// TIA Portal project "PalletWarehouse" (V20)

(* hardware
DEVICE "S7-1500/ET200MP-Station_1"  S7-1500 station
   slot 0: "Profilschiene_0"  Rack  6ES7 590-1***0-0AA0
   slot 1: "PLC_1"  CPU 1513-1 PN  6ES7 513-1AM03-0AB0  V4.0
      slot 3: "CPU-Display_1"  6ES7591-1AA00-0AA0
      slot 32768: "PROFINET-Schnittstelle_1"  X1
         slot 32769: "Port_1"  X1 P1
         slot 32770: "Port_2"  X1 P2
      slot 34817: "Virtual CP interface port_1"  Virtual CP interface port  Virtual CP interface port FW V4.0
   slot 2: "DI 16x24VDC BA_1"  DI 16x24VDC BA  6ES7 521-1BH10-0AA0  V1.1
   slot 3: "DQ 16x24VDC/0.5A ST_1"  DQ 16x24VDC/0.5A ST  6ES7 522-1BH00-0AB0  V2.0
   slot 4: "AI 8xU/I/R/RTD BA_1"  AI 8xU/I/R/RTD BA  6ES7 531-7QF00-0AB0  V1.0
   slot 5: "AQ 8xU/I HS_1"  AQ 8xU/I HS  6ES7 532-5HF00-0AB0  V2.2
   slot 6: "DQ 16x24VDC/0.5A ST_2"  DQ 16x24VDC/0.5A ST  6ES7 522-1BH00-0AB0  V2.0
   slot 7: "DI 16x24VDC BA_2"  DI 16x24VDC BA  6ES7 521-1BH10-0AA0  V1.1
   slot 8: "AQ 2xU/I ST_1"  AQ 2xU/I ST  6ES7 532-5NB00-0AB0  V1.0
   slot 9: "DI 16x24VDC BA_3"  DI 16x24VDC BA  6ES7 521-1BH10-0AA0  V1.1
DEVICE "PC-System_1"  SIMATIC PC station
   slot 0: "SIMATIC PC station"  Rail  SIMATIC PC-Station  V1.0
      slot 125: "Stationmanager"  Station_Manager  V6.0.4
   slot 1: "HMI_RT_1"  WinCC RT Advanced  6AV2 104-0xxxx-xxxx  17.0.0.0
      slot 33792: "Computer interface"  Host interface
   slot 2: "IE general_1"  IE General  IE_CP  V8.2.0
      slot 1: "PROFINET interface"  IEGeneral.Interface.8.2.0
*)

// ===== PLC "PLC_1"  CPU 1513-1 PN =====

VAR_GLOBAL   // PLC tag table "Standard-Variablentabelle"
   "PlcLabConnectIn01" AT %ID32760 : DWord;
   "PlcLabConnectIn02" AT %ID32764 : DWord;
   "PlcLabConnectOut01" AT %QD32760 : DWord;
   "PlcLabConnectOut02" AT %QD32764 : DWord;
END_VAR

VAR_GLOBAL   // PLC tag table "IO"
   "PalletizerEntrySensor" AT %I0.1 : Bool;
   "PusherLimitSensor" AT %I0.3 : Bool;
   "PalletizerBelt" AT %Q0.4 : Bool;
   "PalletizerTurn" AT %Q0.5 : Bool;
   "PusherMotor" AT %Q0.6 : Bool;
   "PalletizerClampedSensor" AT %I0.5 : Bool;
   "PalletizerPlateLimit" AT %I0.4 : Bool;
   "PalletizerElevatorMovingSensor" AT %I0.6 : Bool;
   "PalletizerClamp" AT %Q0.7 : Bool;
   "PalletizerPlate" AT %Q1.0 : Bool;
   "PalletizerElevatorUp" AT %Q1.1 : Bool;
   "PalletizerElevatorDown" AT %Q1.2 : Bool;
   "PalletizerElevatorMoveToLimit" AT %Q1.3 : Bool;
   "BoxEmitter" AT %Q0.1 : Bool;
   "PalletChainFrontLimit" AT %I0.7 : Bool;
   "BoxFeedConveyor" AT %Q0.0 : Bool;
   "PalletChain" AT %Q0.2 : Bool;
   "PalletFeedSensor" AT %I0.2 : Bool;
   "PalletFeedConveyor" AT %Q1.4 : Bool;
   "PalletEmitter" AT %Q0.3 : Bool;
   "ConveyorSensor1" AT %I1.1 : Bool;
   "ConveyorSensor2" AT %I1.2 : Bool;
   "TransferConveyor1" AT %Q1.5 : Bool;
   "TransferConveyor2" AT %Q1.6 : Bool;
   "TurntableEntrySensor" AT %I1.3 : Bool;
   "PalletChainBackLimit" AT %I1.0 : Bool;
   "TurntableTurn" AT %Q1.7 : Bool;
   "TurntableRollForward" AT %Q2.0 : Bool;
   "TurntableRollBackward" AT %Q2.1 : Bool;
   "TurntableLimit0" AT %I1.4 : Bool;
   "TurntableLimit90" AT %I1.5 : Bool;
   "TurntableBackLimit" AT %I1.6 : Bool;
   "TurntableFrontLimit" AT %I1.7 : Bool;
   "TurntableLeftExitSensor" AT %I2.0 : Bool;
   "TurntableRightExitSensor" AT %I2.1 : Bool;
   "Crane1MovingX" AT %I2.2 : Bool;
   "Crane1MovingZ" AT %I2.3 : Bool;
   "Crane1LeftLimit" AT %I2.4 : Bool;
   "Crane1RightLimit" AT %I2.5 : Bool;
   "Crane1Lift" AT %Q2.2 : Bool;
   "Crane1Right" AT %Q2.4 : Bool;
   "Crane1Left" AT %Q2.3 : Bool;
   "Crane1Position" AT %QW30 : Int;
   "StartButtonTemp" AT %I2.7 : Bool;
   "Crane1MidLimit" AT %I2.6 : Bool;
   "Crane2MovingX" AT %I3.0 : Bool;
   "Crane2MovingZ" AT %I3.1 : Bool;
   "Crane2LeftLimit" AT %I3.2 : Bool;
   "Crane2RightLimit" AT %I3.3 : Bool;
   "Crane2MidLimit" AT %I3.4 : Bool;
   "Crane2Lift" AT %Q2.5 : Bool;
   "Crane2Right" AT %Q2.7 : Bool;
   "Crane2Left" AT %Q2.6 : Bool;
   "Crane2Position" AT %QW32 : Int;
   "LoadSensor1" AT %I3.5 : Bool;
   "LoadSensor2" AT %I3.6 : Bool;
   "LoadConveyor1" AT %Q3.0 : Bool;
   "LoadConveyor2" AT %Q3.1 : Bool;
   "BoxEmitterSensor" AT %I0.0 : Bool;
   "UnloadSensor1" AT %I3.7 : Bool;
   "UnloadSensor2" AT %I4.0 : Bool;
   "RemoverSensor1" AT %I4.1 : Bool;
   "RemoverSensor2" AT %I4.2 : Bool;
   "UnloadConveyor1" AT %Q3.2 : Bool;
   "UnloadConveyor2" AT %Q3.3 : Bool;
   "RemoverConveyor1" AT %Q3.4 : Bool;
   "RemoverConveyor2" AT %Q3.5 : Bool;
   "Remover1" AT %Q3.6 : Bool;
   "Remover2" AT %Q3.7 : Bool;
END_VAR

TYPE "StorageCraneUDT"
   STRUCT
      CraneSides : Struct
         LoadRight : Bool;
         UnloadRight : Bool;
         PickupRight : Bool;
      END_STRUCT;
      In : Struct
         MovingX : Bool;
         MovingZ : Bool;
         LeftLimit : Bool;
         RightLimit : Bool;
         MidLimit : Bool;
      END_STRUCT;
      Out : Struct
         Lift : Bool;
         Left : Bool;
         Right : Bool;
         Position : Int;
      END_STRUCT;
   END_STRUCT;
END_TYPE

TYPE "WarehouseSlotUDT"
   STRUCT
      Id : Int;
      Status : Int;
      "Time" : DTL;
   END_STRUCT;
END_TYPE

TYPE "PalletizerUDT"
   STRUCT
      In : Struct
         BoxEntrySensor : Bool;
         PusherLimit : Bool;
         Clamped : Bool;
         PlateLimit : Bool;
         ElevatorMoving : Bool;
         ElevatorFrontLimit : Bool;
         ElevatorBackLimit : Bool;
         PalletFeedSensor : Bool;
         EmitSensor : Bool;
      END_STRUCT;
      Out : Struct
         PalletFeedConv : Bool;
         BoxFeedConv : Bool;
         Turn : Bool;
         Clamp : Bool;
         Pusher : Bool;
         Plate : Bool;
         ElevatorUp : Bool;
         ElevatorDown : Bool;
         ElevatorMoveToLimit : Bool;
         PalletConv : Bool;
         PalletEmitter : Bool;
         EmitConv : Bool;
         BoxEmitter : Bool;
      END_STRUCT;
   END_STRUCT;
END_TYPE

TYPE "ConveyorUDT"
   STRUCT
      In : Struct
         StartSensor : Bool;
         EndSensor : Bool;
         Stop : Bool;
      END_STRUCT;
      Out : Struct
         Conveyor : Bool;
      END_STRUCT;
   END_STRUCT;
END_TYPE

TYPE "TurntableUDT"
   STRUCT
      In : Struct
         FrontLimit : Bool;
         BackLimit : Bool;
         Limit90 : Bool;
         Limit0 : Bool;
      END_STRUCT;
      Out : Struct
         RollForward : Bool;
         RollBackward : Bool;
         Turn : Bool;
      END_STRUCT;
   END_STRUCT;
END_TYPE

DATA_BLOCK "Warehouse_DB"   // DB9
{ S7_Optimized_Access := 'TRUE' }
VERSION : 0.1
// stored: InstanceOfName Warehouse
"Warehouse"
BEGIN
END_DATA_BLOCK

// folder: HMI

DATA_BLOCK "HMI_Data"   // DB11
{ S7_Optimized_Access := 'TRUE' }
VERSION : 0.1
   VAR
      SelectedRack : Int;
      SelectedSlot : Int;
      TargetSlot : "WarehouseSlotUDT";
      RetrievePallet : Bool;
      StopCmd : Bool;
      StartCmd : Bool;
      RacksFull : Bool;
      CraneStatus : Array[1..2] of Int;
      OccupiedSlots : Array[1..2] of Int;
   END_VAR
BEGIN
END_DATA_BLOCK

// folder: IO Mapping

DATA_BLOCK "IO"   // DB2
{ S7_Optimized_Access := 'TRUE' }
VERSION : 0.1
   VAR
      Palletizer : "PalletizerUDT";
      StorageCrane1 : "StorageCraneUDT";
      StorageCrane2 : "StorageCraneUDT";
      LineIO : Struct
         TransferConveyor1IO : "ConveyorUDT";
         TransferConveyor2IO : "ConveyorUDT";
         LoadConveyor1IO : "ConveyorUDT";
         LoadConveyor2IO : "ConveyorUDT";
         UnloadConveyor1IO : "ConveyorUDT";
         UnloadConveyor2IO : "ConveyorUDT";
         TurntableIO : "TurntableUDT";
         Remover1 : Bool;
         Remover2 : Bool;
      END_STRUCT;
   END_VAR
BEGIN
   StorageCrane1.CraneSides.LoadRight := TRUE;
   StorageCrane1.CraneSides.PickupRight := TRUE;
   StorageCrane1.CraneSides.UnloadRight := FALSE;
   StorageCrane2.CraneSides.PickupRight := FALSE;
   StorageCrane2.CraneSides.UnloadRight := TRUE;
   StorageCrane2.CraneSides.LoadRight := TRUE;
END_DATA_BLOCK

// folder: WarehouseManager

DATA_BLOCK "WarehouseData"   // DB10
{ S7_Optimized_Access := 'TRUE' }
VERSION : 0.1
   VAR
      Rack1 : Array[1..54] of "WarehouseSlotUDT";
      Rack2 : Array[1..54] of "WarehouseSlotUDT";
   END_VAR
BEGIN
END_DATA_BLOCK

// folder: (top level)

FUNCTION_BLOCK "Warehouse"   // FB15, SCL
{ S7_Optimized_Access := 'TRUE' }
VERSION : 0.1
   VAR_IN_OUT
      PalletizerIO : "PalletizerUDT";
      StorageCrane1IO : "StorageCraneUDT";
      StorageCrane2IO : "StorageCraneUDT";
      LineIO : Struct
         TransferConveyor1IO : "ConveyorUDT";
         TransferConveyor2IO : "ConveyorUDT";
         LoadConveyor1IO : "ConveyorUDT";
         LoadConveyor2IO : "ConveyorUDT";
         UnloadConveyor1IO : "ConveyorUDT";
         UnloadConveyor2IO : "ConveyorUDT";
         TurntableIO : "TurntableUDT";
         Remover1 : Bool;
         Remover2 : Bool;
      END_STRUCT;
   END_VAR
   VAR
      Line : "Line";
      WarehouseManager : "WarehouseManager";
      CraneLoadDone : Array[1..2] of Bool;
      CraneUnloadDone : Array[1..2] of Bool;
      CraneBusy : Array[1..2] of Bool;
      Palletizer : "Palletizer";
      StorageCrane1 : "StorageCrane";
      StorageCrane2 : "StorageCrane";
      WarehouseControl : "WarehouseControl";
   END_VAR
BEGIN
   #WarehouseControl(StartCmd := "HMI_Data".StartCmd,
                     StopCmd := "HMI_Data".StopCmd,
                     Active := false);

   #Palletizer(PalletizerIO:=#PalletizerIO,
               Run:=#WarehouseControl.Run AND NOT #WarehouseManager.Full);

   #WarehouseManager(UnloadDone:=#CraneUnloadDone,
                     CraneBusy:=#CraneBusy,
                     PalletReady := #LineIO.TransferConveyor2IO.In.EndSensor,
                     UnloadRequest:="HMI_Data".RetrievePallet,
                     UnloadRack:="HMI_Data".SelectedRack,
                     UnloadSlot:="HMI_Data".SelectedSlot,
                     Run:=#WarehouseControl.Run,
                     Rack1Slots := "WarehouseData".Rack1,
                     Rack2Slots := "WarehouseData".Rack2,
                     LoadDone:=#CraneLoadDone,
                     Full=>"HMI_Data".RacksFull,
                     CraneStatus=>"HMI_Data".CraneStatus); 

   #Line(TurntableRollDirection:=#WarehouseManager.Rack,
         Run:=#WarehouseControl.Run,
         Remover1=>#LineIO.Remover1,
         Remover2=>#LineIO.Remover2,
         TransferConveyor1IO:=#LineIO.TransferConveyor1IO,
         TransferConveyor2IO:=#LineIO.TransferConveyor2IO,
         LoadConveyor1IO:=#LineIO.LoadConveyor1IO,
         LoadConveyor2IO:=#LineIO.LoadConveyor2IO,
         UnloadConveyor1IO:=#LineIO.UnloadConveyor1IO,
         UnloadConveyor2IO:=#LineIO.UnloadConveyor2IO,
         TurntableIO:=#LineIO.TurntableIO);

   #StorageCrane1(TargetPosition:=#WarehouseManager.TargetSlot[1],
                  RequestLoad:=#WarehouseManager.LoadStart[1] AND #LineIO.LoadConveyor1IO.In.Stop,
                  RequestUnload:=#WarehouseManager.UnloadStart[1],
                  Run:=#WarehouseControl.Run,
                  LoadDone=>#CraneLoadDone[1],
                  UnloadDone=>#CraneUnloadDone[1],
                  StorageCraneUDT:=#StorageCrane1IO,
                  Busy=>#CraneBusy[1]); 

   #StorageCrane2(TargetPosition := #WarehouseManager.TargetSlot[2],
                  RequestLoad := #WarehouseManager.LoadStart[2] AND #LineIO.LoadConveyor2IO.In.Stop,
                  RequestUnload := #WarehouseManager.UnloadStart[2],
                  Run:=#WarehouseControl.Run,
                  LoadDone => #CraneLoadDone[2],
                  UnloadDone=>#CraneUnloadDone[2],
                  StorageCraneUDT := #StorageCrane2IO,
                  Busy=>#CraneBusy[2]);
END_FUNCTION_BLOCK

FUNCTION_BLOCK "WarehouseControl"   // FB19, SCL
{ S7_Optimized_Access := 'TRUE' }
VERSION : 0.1
   VAR_INPUT
      StartCmd : Bool;
      StopCmd : Bool;
      Active : Bool;
   END_VAR
   VAR_OUTPUT
      Run : Bool;
      Status : Int;
   END_VAR
   VAR
      StopPEdge : R_TRIG;
      StartPEdge : R_TRIG;
   END_VAR
BEGIN
   #StartPEdge(CLK:=#StartCmd);
   #StopPEdge(CLK := #StopCmd);

   IF #StopPEdge.Q THEN
       #Run := FALSE;
   ELSIF #StartPEdge.Q THEN
       #Run := TRUE;
   END_IF;

   IF #Run THEN
       #Status := 1;
   ELSIF #Active THEN
       #Status := 2;
   ELSE
       #Status := 0;
   END_IF;
END_FUNCTION_BLOCK

ORGANIZATION_BLOCK "Main"   // OB1, LAD, ProgramCycle
TITLE = "Main Program Sweep (Cycle)"
{ S7_Optimized_Access := 'TRUE' }
VERSION : 0.1
   VAR_INPUT
      Initial_Call : Bool;   // Initial call of this OB
      Remanence : Bool;   // =True, if remanent data are available
   END_VAR
BEGIN

REGION Network 1
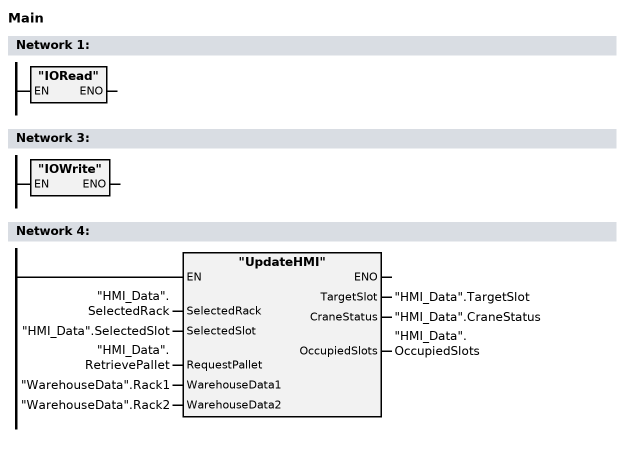
   RUNG wire#powerrail
      "IORead"()
   END_RUNG
   // the same network as SCL:
   "IORead"();
END_REGION

REGION Network 2 (SCL)
   "Warehouse_DB"(PalletizerIO:="IO".Palletizer,
                  StorageCrane1IO:="IO".StorageCrane1,
                  StorageCrane2IO:="IO".StorageCrane2,
                  LineIO:="IO".LineIO);
END_REGION

REGION Network 3
   RUNG wire#powerrail
      "IOWrite"()
   END_RUNG
   // the same network as SCL:
   "IOWrite"();
END_REGION

REGION Network 4
   RUNG wire#powerrail
      "UpdateHMI"(SelectedRack := "HMI_Data".SelectedRack, SelectedSlot := "HMI_Data".SelectedSlot, RequestPallet := "HMI_Data".RetrievePallet, WarehouseData1 := "WarehouseData".Rack1, WarehouseData2 := "WarehouseData".Rack2, TargetSlot => "HMI_Data".TargetSlot, CraneStatus => "HMI_Data".CraneStatus, OccupiedSlots => "HMI_Data".OccupiedSlots)
   END_RUNG
   // the same network as SCL:
   "UpdateHMI"(SelectedRack := "HMI_Data".SelectedRack,
               SelectedSlot := "HMI_Data".SelectedSlot,
               RequestPallet := "HMI_Data".RetrievePallet,
               WarehouseData1 := "WarehouseData".Rack1,
               WarehouseData2 := "WarehouseData".Rack2,
               TargetSlot => "HMI_Data".TargetSlot,
               CraneStatus => "HMI_Data".CraneStatus,
               OccupiedSlots => "HMI_Data".OccupiedSlots);
END_REGION
END_ORGANIZATION_BLOCK

// folder: HMI

FUNCTION "UpdateHMI" : Void   // FC6, SCL
{ S7_Optimized_Access := 'TRUE' }
VERSION : 0.1
   VAR_INPUT
      SelectedRack : Int;
      SelectedSlot : Int;
      RequestPallet : Bool;
      WarehouseData1 : Array[1..54] of "WarehouseSlotUDT";
      WarehouseData2 : Array[1..54] of "WarehouseSlotUDT";
   END_VAR
   VAR_OUTPUT
      TargetSlot : "WarehouseSlotUDT";
      CraneStatus : Array[1..2] of Int;
      OccupiedSlots : Array[1..2] of Int;
   END_VAR
   VAR_TEMP
      i : Int;
      freeslots : Array[1..2] of Int;
   END_VAR
BEGIN
   IF #SelectedRack = 1 THEN
       #TargetSlot := #WarehouseData1[#SelectedSlot];
   ELSIF #SelectedRack = 2 THEN
       #TargetSlot := #WarehouseData2[#SelectedSlot];
   END_IF;

   #freeslots[1]:="CountFreeSlots"(#WarehouseData1);
   #freeslots[2] := "CountFreeSlots"(#WarehouseData2);

   FOR #i := 1 TO 2 DO
       #OccupiedSlots[#i] := 54 - #freeslots[#i];
   END_FOR;
END_FUNCTION

// folder: IO Mapping

FUNCTION "IOWrite" : Void   // FC4, SCL
{ S7_Optimized_Access := 'TRUE' }
VERSION : 0.1
BEGIN
   // Mapping palletizer outputs
   "PalletFeedConveyor":="IO".Palletizer.Out.PalletFeedConv;
   "PalletizerBelt" :="IO".Palletizer.Out.BoxFeedConv;
   "PalletizerTurn" :="IO".Palletizer.Out.Turn;
   "PalletizerClamp":="IO".Palletizer.Out.Clamp;
   "PusherMotor" :="IO".Palletizer.Out.Pusher;
   "PalletizerPlate" := "IO".Palletizer.Out.Plate;
   "PalletizerElevatorUp" := "IO".Palletizer.Out.ElevatorUp;
   "PalletizerElevatorDown" :="IO".Palletizer.Out.ElevatorDown;
   "PalletizerElevatorMoveToLimit" :="IO".Palletizer.Out.ElevatorMoveToLimit;
   "PalletChain":="IO".Palletizer.Out.PalletConv;
   "PalletEmitter":="IO".Palletizer.Out.PalletEmitter;
   "BoxEmitter" := "IO".Palletizer.Out.BoxEmitter;
   "BoxFeedConveyor" := "IO".Palletizer.Out.EmitConv;

   // Mapping storage crane 1 outputs
   "Crane1Lift" := "IO".StorageCrane1.Out.Lift;
   "Crane1Left" :="IO".StorageCrane1.Out.Left;
   "Crane1Right" := "IO".StorageCrane1.Out.Right;
   "Crane1Position" := "IO".StorageCrane1.Out.Position;
   // Mapping storage crane 2 outputs
   "Crane2Lift":="IO".StorageCrane2.Out.Lift;
   "Crane2Left":="IO".StorageCrane2.Out.Left;
   "Crane2Right":="IO".StorageCrane2.Out.Right;
   "Crane2Position" := "IO".StorageCrane2.Out.Position;
   // Mapping line outputs
   "TransferConveyor1":="IO".LineIO.TransferConveyor1IO.Out.Conveyor;
   "TransferConveyor2":="IO".LineIO.TransferConveyor2IO.Out.Conveyor;
   "TurntableRollForward" := "IO".LineIO.TurntableIO.Out.RollForward;
   "TurntableRollBackward" := "IO".LineIO.TurntableIO.Out.RollBackward;
   "TurntableTurn" := "IO".LineIO.TurntableIO.Out.Turn;
   "LoadConveyor1":="IO".LineIO.LoadConveyor1IO.Out.Conveyor;
   "LoadConveyor2":="IO".LineIO.LoadConveyor2IO.Out.Conveyor;
   "UnloadConveyor1" := "IO".LineIO.UnloadConveyor1IO.Out.Conveyor;
   "UnloadConveyor2" := "IO".LineIO.UnloadConveyor2IO.Out.Conveyor;
   "RemoverConveyor1" := "IO".LineIO.UnloadConveyor1IO.Out.Conveyor;
   "RemoverConveyor2" := "IO".LineIO.UnloadConveyor2IO.Out.Conveyor;
   "Remover1" := "IO".LineIO.Remover1;
   "Remover2" := "IO".LineIO.Remover2;
END_FUNCTION

FUNCTION "IORead" : Void   // FC5, SCL
{ S7_Optimized_Access := 'TRUE' }
VERSION : 0.1
BEGIN
   // Mapping Palletizer Inputs
   "IO".Palletizer.In.BoxEntrySensor := "PalletizerEntrySensor";
   "IO".Palletizer.In.PusherLimit := "PusherLimitSensor";
   "IO".Palletizer.In.Clamped := "PalletizerClampedSensor";
   "IO".Palletizer.In.PlateLimit := "PalletizerPlateLimit";
   "IO".Palletizer.In.ElevatorMoving := "PalletizerElevatorMovingSensor";
   "IO".Palletizer.In.ElevatorFrontLimit := "PalletChainFrontLimit";
   "IO".Palletizer.In.ElevatorBackLimit := "PalletChainBackLimit";
   "IO".Palletizer.In.PalletFeedSensor := "PalletFeedSensor";
   "IO".Palletizer.In.EmitSensor := "BoxEmitterSensor";
   // Maping Storage Crane 1 Inputs
   "IO".StorageCrane1.In.MovingX := "Crane1MovingX";
   "IO".StorageCrane1.In.MovingZ := "Crane1MovingZ";
   "IO".StorageCrane1.In.LeftLimit := "Crane1LeftLimit";
   "IO".StorageCrane1.In.RightLimit := "Crane1RightLimit";
   "IO".StorageCrane1.In.MidLimit := "Crane1MidLimit";
   // Maping Storage Crane 2 Inputs
   "IO".StorageCrane2.In.MovingX := "Crane2MovingX";
   "IO".StorageCrane2.In.MovingZ := "Crane2MovingZ";
   "IO".StorageCrane2.In.LeftLimit := "Crane2LeftLimit";
   "IO".StorageCrane2.In.RightLimit := "Crane2RightLimit";
   "IO".StorageCrane2.In.MidLimit := "Crane2MidLimit";
   // Maping Line Inputs
   "IO".LineIO.TransferConveyor1IO.In.StartSensor := "ConveyorSensor1";
   "IO".LineIO.TransferConveyor1IO.In.EndSensor := "ConveyorSensor2";
   "IO".LineIO.TransferConveyor2IO.In.StartSensor := "ConveyorSensor2";
   "IO".LineIO.TransferConveyor2IO.In.EndSensor := "TurntableEntrySensor";
   "IO".LineIO.TurntableIO.In.FrontLimit := "TurntableFrontLimit";
   "IO".LineIO.TurntableIO.In.BackLimit := "TurntableBackLimit";
   "IO".LineIO.TurntableIO.In.Limit90 := "TurntableLimit90";
   "IO".LineIO.TurntableIO.In.Limit0 := "TurntableLimit0";
   "IO".LineIO.LoadConveyor1IO.In.StartSensor := "TurntableLeftExitSensor";
   "IO".LineIO.LoadConveyor1IO.In.Stop := "LoadSensor1";
   "IO".LineIO.LoadConveyor2IO.In.StartSensor := "TurntableRightExitSensor";
   "IO".LineIO.LoadConveyor2IO.In.Stop := "LoadSensor2";
   "IO".LineIO.UnloadConveyor1IO.In.StartSensor := "UnloadSensor1";
   "IO".LineIO.UnloadConveyor2IO.In.StartSensor := "UnloadSensor2";
   "IO".LineIO.UnloadConveyor1IO.In.Stop := "RemoverSensor1";
   "IO".LineIO.UnloadConveyor2IO.In.Stop := "RemoverSensor2";
END_FUNCTION

// folder: Line

FUNCTION_BLOCK "Line"   // FB1, LAD
{ S7_Optimized_Access := 'TRUE' }
VERSION : 0.1
   VAR_INPUT
      TurntableRollDirection : Int;
      Run : Bool;
   END_VAR
   VAR_OUTPUT
      Remover1 : Bool;
      Remover2 : Bool;
   END_VAR
   VAR_IN_OUT
      TransferConveyor1IO : "ConveyorUDT";
      TransferConveyor2IO : "ConveyorUDT";
      LoadConveyor1IO : "ConveyorUDT";
      LoadConveyor2IO : "ConveyorUDT";
      UnloadConveyor1IO : "ConveyorUDT";
      UnloadConveyor2IO : "ConveyorUDT";
      TurntableIO : "TurntableUDT";
   END_VAR
   VAR
      UnloadConveyor2 : "Conveyor";
      TransferConveyor1 : "Conveyor";
      TransferConveyor2 : "Conveyor";
      Turntable : "Turntable";
      LoadConveyor1 : "Conveyor";
      LoadConveyor2 : "Conveyor";
      UnloadConveyor1 : "Conveyor";
   END_VAR
BEGIN

REGION Network 1 (SCL)
   #TransferConveyor1(NextFree:=NOT #TransferConveyor2.Busy,
                      Run:=#Run,
                      ConveyorIO:=#TransferConveyor1IO);  

   #TransferConveyor2(NextFree:=TRUE,
                      Run:=#Run,
                      ConveyorIO:=#TransferConveyor2IO);

   #Turntable(Start:=#TransferConveyor2IO.In.EndSensor,
              Run:=#Run,
              RollDirection:=#TurntableRollDirection,
              RightSensor:=#LoadConveyor2IO.In.StartSensor,
              LeftSensor:=#LoadConveyor1IO.In.StartSensor,
              TurntableIO:=#TurntableIO); 

   #LoadConveyor1(NextFree:=TRUE,
                  Run:=#Run,
                  ConveyorIO:=#LoadConveyor1IO);

   #LoadConveyor2(NextFree:=TRUE,
                  Run:=#Run,
                  ConveyorIO:=#LoadConveyor2IO);

   #UnloadConveyor1(NextFree:=TRUE,
                    Run:=#Run,
                    ConveyorIO:=#UnloadConveyor1IO);

   #UnloadConveyor2(NextFree:=TRUE,
                    Run:=#Run,
                    ConveyorIO:=#UnloadConveyor2IO);

   #Remover1 := #UnloadConveyor1IO.In.Stop;
   #Remover2 := #UnloadConveyor2IO.In.Stop;
END_REGION
END_FUNCTION_BLOCK

FUNCTION_BLOCK "Conveyor"   // FB2, LAD
{ S7_Optimized_Access := 'TRUE' }
VERSION : 0.1
   VAR_INPUT
      NextFree : Bool;
      Run : Bool;
   END_VAR
   VAR_OUTPUT
      Busy : Bool;
   END_VAR
   VAR_IN_OUT
      ConveyorIO : "ConveyorUDT";
   END_VAR
   VAR
      Reset : Bool;
      Timeout_Instance : TON_TIME;
      Timeout : Bool;
      StartSensorEdge : Bool;
      EndSensorEdge : Bool;
      ConveyorStart : Bool;
   END_VAR
   VAR_TEMP   // added for the SCL form of the ladder/FBD networks
      _w1 : Bool;
   END_VAR
BEGIN

REGION Network 1
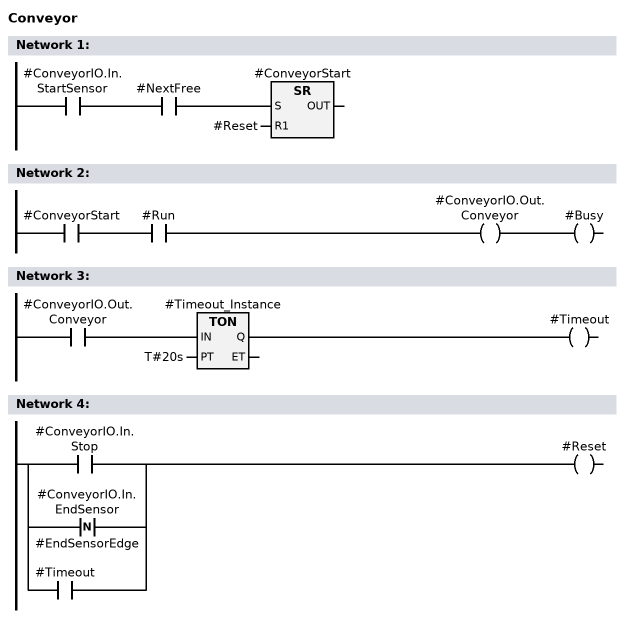
   RUNG wire#powerrail
      Contact( #ConveyorIO.In.StartSensor )
      Contact( #NextFree )
      S_SR(operand := #ConveyorStart, r1 := #Reset)
   END_RUNG
   // the same network as SCL:
   IF #ConveyorIO.In.StartSensor AND #NextFree THEN
       #ConveyorStart := TRUE;   // SR flip-flop
   END_IF;
   IF #Reset THEN #ConveyorStart := FALSE; END_IF;
END_REGION

REGION Network 2
   RUNG wire#powerrail
      Contact( #ConveyorStart )
      Contact( #Run )
      Coil( #ConveyorIO.Out.Conveyor )
      Coil( #Busy )
   END_RUNG
   // the same network as SCL:
   #ConveyorIO.Out.Conveyor := #ConveyorStart AND #Run;
   #Busy := #ConveyorIO.Out.Conveyor;
END_REGION

REGION Network 3
   #Timeout_Instance(IN := #ConveyorIO.Out.Conveyor, PT := T#20s);   // TON
   #Timeout := #Timeout_Instance.Q;
END_REGION

REGION Network 4
   RUNG wire#powerrail
      Contact( #ConveyorIO.In.Stop )
      wire#w1
      Coil( #Reset )
   END_RUNG
   RUNG wire#powerrail
      N_Contact(operand := #ConveyorIO.In.EndSensor, bit := #EndSensorEdge)
   END_RUNG wire#w1
   RUNG wire#powerrail
      Contact( #Timeout )
   END_RUNG wire#w1
   // the same network as SCL:
   #_w1 := NOT #ConveyorIO.In.EndSensor AND #EndSensorEdge;   // falling edge of #ConveyorIO.In.EndSensor
   #EndSensorEdge := #ConveyorIO.In.EndSensor;
   #Reset := #ConveyorIO.In.Stop OR #_w1 OR #Timeout;
END_REGION
END_FUNCTION_BLOCK

FUNCTION_BLOCK "Turntable"   // FB7, SCL
{ S7_Optimized_Access := 'TRUE' }
VERSION : 0.1
   VAR_INPUT
      Start : Bool;
      Run : Bool;
      RollDirection : Int;
      RightSensor : Bool;
      LeftSensor : Bool;
   END_VAR
   VAR_IN_OUT
      TurntableIO : "TurntableUDT";
   END_VAR
   VAR
      State : Int := 1;
      RightSensorNEdge : F_TRIG;
      LeftSensorNEdge : F_TRIG;
   END_VAR
BEGIN
   #RightSensorNEdge(CLK:=#RightSensor);
   #LeftSensorNEdge(CLK:=#LeftSensor);

   CASE #State OF
       1:  // Init
           IF #Start THEN
               #State := 2;
           END_IF;
           ;
       2:  // Load
           "IO".LineIO.TurntableIO.Out.RollForward := #Run;
           IF #TurntableIO.In.FrontLimit THEN
               #TurntableIO.Out.RollForward := FALSE;
               #State := 3;
           END_IF;
           ;
       3: // Turn
           #TurntableIO.Out.Turn := TRUE;
           IF #TurntableIO.In.Limit90 THEN
               #State := 4;
           END_IF;
       4: // Direction
           IF #RollDirection=1 THEN
               #State := 5;
           ELSIF #RollDirection=2 THEN
               #State := 6;
           END_IF;
       5: // Roll left
           #TurntableIO.Out.RollForward := #Run;
           IF #LeftSensorNEdge.Q THEN
               #TurntableIO.Out.RollForward := FALSE;
               #State := 7;
           END_IF;
       6: // Roll right
           #TurntableIO.Out.RollBackward := #Run;
           IF #RightSensorNEdge.Q THEN
               #TurntableIO.Out.RollBackward := FALSE;
               #State := 7;
           END_IF;
       7: // Return 
           #TurntableIO.Out.Turn := FALSE;
           IF #TurntableIO.In.Limit0 THEN
               #State := 1;
           END_IF;
   END_CASE;
END_FUNCTION_BLOCK

// folder: Palletizer

FUNCTION_BLOCK "Palletizer"   // FB3, SCL
{ S7_Optimized_Access := 'TRUE' }
VERSION : 0.1
   VAR_INPUT
      Run : Bool;
   END_VAR
   VAR_OUTPUT
      Busy : Bool;
   END_VAR
   VAR_IN_OUT
      PalletizerIO : "PalletizerUDT";
   END_VAR
   VAR
      State : Int := 1;
      BoxCount : Int := 0;
      BoxFeedTimer : TON_TIME;
      BoxFeedBusy : Bool;
      StackVertical : Bool := TRUE;
      PushCount : Int;
      BoxEntrySensorNEdge : F_TRIG;
      PusherFB : "Cylinder";
      BoxPerPush : Int;
      PushPerLayer : Int;
      PlateFB : "Cylinder";
      ElevatorFB : "Elevator";
      LayerCount : Int;
      PalletFeederFB : "PalletFeeder";
      BoxFeeder : "BoxFeedConv";
      UnloadConv : Bool;
   END_VAR
BEGIN
   #BoxEntrySensorNEdge(CLK := #PalletizerIO.In.BoxEntrySensor);
   #BoxFeedTimer(IN:=#PalletizerIO.Out.BoxFeedConv AND #BoxCount=#BoxPerPush,
                 PT:=T#2s);

   #PusherFB.Extend := FALSE;
   #PlateFB.Extend := FALSE;
   #PalletizerIO.Out.Clamp := FALSE;
   #PalletizerIO.Out.PalletConv := FALSE;
   #PalletFeederFB.Start := FALSE;
   #ElevatorFB.RequestUp := FALSE;
   #ElevatorFB.RequestDown := FALSE;
   #ElevatorFB.GoToLimit := FALSE;
   #UnloadConv := FALSE;

   IF #BoxEntrySensorNEdge.Q THEN
       #BoxCount := #BoxCount + 1;
   END_IF;

   IF #StackVertical THEN
       #PalletizerIO.Out.Turn := FALSE;
       #BoxPerPush := 2;
       #PushPerLayer := 3;
   ELSE
       #PalletizerIO.Out.Turn := TRUE;
       #BoxPerPush := 3;
       #PushPerLayer := 2;
   END_IF;

   CASE #State OF
       1:  // Init
           #StackVertical := True;
           #PushCount := 0;
           #BoxCount := 0;
           #LayerCount := 0;
           IF #Run THEN
               #State := 2;
           END_IF;
       2: // Pallet feed
           #PalletFeederFB.Start := #Run;
           IF #PalletFeederFB.Done THEN
               #State := 3;
           END_IF;

       3: // Elevator ready
           #ElevatorFB.GoToLimit := TRUE;
           #ElevatorFB.RequestUp := TRUE;
           IF #ElevatorFB.Done THEN
               #State := 4;
           END_IF;

       4:  // Box feed
           IF #PalletizerIO.In.BoxEntrySensor AND (#BoxCount < #BoxPerPush) AND #Run THEN
               #PalletizerIO.Out.BoxFeedConv := TRUE;
           ELSIF #BoxFeedTimer.Q THEN
               #PalletizerIO.Out.BoxFeedConv := FALSE;
           ELSIF (#BoxCount<#BoxPerPush) AND (NOT #Run) THEN
               #PalletizerIO.Out.BoxFeedConv := FALSE;
           END_IF;

           IF #BoxCount = #BoxPerPush AND NOT #PalletizerIO.Out.BoxFeedConv THEN
               #BoxCount := 0;
               #State := 5;
           END_IF;

       5:  // Extend pusher
           #PusherFB.Extend := TRUE;
           IF #PusherFB.Extended THEN
               #PushCount := #PushCount + 1;
               #State := 6;
           END_IF;

       6:  // Retract pusher
           IF #PusherFB.Retracted THEN
               IF #PushCount >= #PushPerLayer THEN
                   #PushCount := 0;
                   #StackVertical := NOT #StackVertical;
                   #State := 7;
               ELSE
                   #State := 4;
               END_IF;
           END_IF;

       7:  // Clamp
           #PalletizerIO.Out.Clamp := TRUE;
           IF #PalletizerIO.In.Clamped THEN
               #State := 8;
           END_IF;

       8: // Plate open
           #PalletizerIO.Out.Clamp := TRUE;
           #PlateFB.Extend := TRUE;
           IF #PlateFB.Extended THEN
               #State := 9;
           END_IF;

       9: // Layer down
           #ElevatorFB.RequestDown := TRUE;
           #PlateFB.Extend := TRUE;
           IF #ElevatorFB.Done THEN
               #LayerCount := #LayerCount + 1;
               #State := 10;
           END_IF;

       10: // Plate close
           IF #PlateFB.Retracted THEN
               #State := 11;
           END_IF;

       11: // Layer check
           IF #LayerCount = 3 THEN
               #State := 12;
           ELSE
               #State := 4;
           END_IF;

       12: // Elevator down
           #ElevatorFB.RequestDown := TRUE;
           #ElevatorFB.GoToLimit := TRUE;
           IF #ElevatorFB.Done THEN
               #State := 13;
           END_IF;
       13: // Unload pallet
           #UnloadConv := #Run;
           IF NOT #PalletizerIO.In.ElevatorFrontLimit THEN
               #State := 1;
           END_IF;
   END_CASE;

   #Busy := (#BoxCount = #BoxPerPush) OR (#State <> 4);

   #PusherFB(LimitSensor := #PalletizerIO.In.PusherLimit,
             Cylinder => #PalletizerIO.Out.Pusher);
   #PlateFB(LimitSensor := #PalletizerIO.In.PlateLimit,
            Cylinder => #PalletizerIO.Out.Plate);
   #ElevatorFB(MovingSensor := #PalletizerIO.In.ElevatorMoving,
               ElevatorUp => #PalletizerIO.Out.ElevatorUp,
               ElevatorDown => #PalletizerIO.Out.ElevatorDown,
               MoveToLimit => #PalletizerIO.Out.ElevatorMoveToLimit);
   #PalletFeederFB(ElevatorFrontLimit := #PalletizerIO.In.ElevatorFrontLimit,
                   PalletSensor := #PalletizerIO.In.PalletFeedSensor,
                   PalletEmitter => #PalletizerIO.Out.PalletEmitter,
                   PalletConveyor => #PalletizerIO.Out.PalletFeedConv);
   #BoxFeeder(Run:=#Run,
              BoxCount := #BoxCount,
              StopCount := #BoxPerPush,
              EndSensor := #PalletizerIO.In.BoxEntrySensor,
              NextBusy := #Busy,
              BoxEmitter => #PalletizerIO.Out.BoxEmitter,
              Conveyor => #PalletizerIO.Out.EmitConv,
              EmitSensor := #PalletizerIO.In.EmitSensor);

   #PalletizerIO.Out.PalletConv := #UnloadConv OR #PalletFeederFB.ElevatorConveyor;
END_FUNCTION_BLOCK

FUNCTION_BLOCK "Cylinder"   // FB4, SCL
{ S7_Optimized_Access := 'TRUE' }
VERSION : 0.1
   VAR_INPUT
      LimitSensor : Bool;
      Extend : Bool;
   END_VAR
   VAR_OUTPUT
      Cylinder : Bool;
      Extended : Bool;
      Retracted : Bool;
   END_VAR
   VAR
      State : Int := 1;
      LastPosition : Bool;
      LeftLimit : Bool;
   END_VAR
BEGIN
   CASE #State OF
       1:  // Init
           #LastPosition := FALSE;
           IF NOT #Extend AND #LimitSensor THEN
               #State := 2;
           ELSE
               #LeftLimit := NOT #LimitSensor;
               #State := 3;
           END_IF;
       2:  // Settled
           IF #Extend <> #LastPosition THEN
               #LeftLimit := FALSE;
               #State := 3;
           END_IF;
       3:  // Moving
           IF NOT #LimitSensor THEN
               #LeftLimit := TRUE;
           END_IF;

           IF #LeftLimit AND #LimitSensor THEN
               #LastPosition := #Extend;
               #State := 2;
           ELSIF NOT #LeftLimit AND (#Extend = #LastPosition) THEN
               #State := 2;
           END_IF;
           ;
   END_CASE;

   #Cylinder := #Extend;
   #Extended := (#State = 2) AND #LastPosition;
   #Retracted := (#State = 2) AND NOT #LastPosition;
END_FUNCTION_BLOCK

FUNCTION_BLOCK "Elevator"   // FB5, SCL
{ S7_Optimized_Access := 'TRUE' }
VERSION : 0.1
   VAR_INPUT
      RequestUp : Bool;
      RequestDown : Bool;
      GoToLimit : Bool;
      MovingSensor : Bool;
   END_VAR
   VAR_OUTPUT
      ElevatorUp : Bool;
      ElevatorDown : Bool;
      Done : Bool;
      MoveToLimit : Bool;
   END_VAR
   VAR
      State : Int := 1;
      RequestUpPEdge : R_TRIG;
      RequestDownPEdge : R_TRIG;
   END_VAR
BEGIN
   #Done := FALSE;
   #RequestUpPEdge(CLK:=#RequestUp);
   #RequestDownPEdge(CLK:=#RequestDown);


   CASE #State OF
       1:  // Idle
           #MoveToLimit := #GoToLimit;
           IF #RequestUpPEdge.Q AND NOT #RequestDown THEN
               #ElevatorUp := TRUE;
               #State := 2;
           ELSIF #RequestDownPEdge.Q AND NOT #RequestUp THEN
               #ElevatorDown := TRUE;
               #State := 2;
           END_IF;
           ;
       2:  // WaitStart
           IF #MovingSensor THEN
               #State := 3;
           END_IF;
           ;
       3: // Moving
           IF NOT #MovingSensor THEN
               #Done := TRUE;
               #ElevatorDown := FALSE;
               #ElevatorUp := FALSE;
               #State := 1;
           END_IF;
           ;
   END_CASE;
END_FUNCTION_BLOCK

FUNCTION_BLOCK "PalletFeeder"   // FB6, SCL
{ S7_Optimized_Access := 'TRUE' }
VERSION : 0.1
   VAR_INPUT
      ElevatorFrontLimit : Bool;
      PalletSensor : Bool;
      Start : Bool;
   END_VAR
   VAR_OUTPUT
      PalletEmitter : Bool;
      PalletConveyor : Bool;
      ElevatorConveyor : Bool;
      Done : Bool;
   END_VAR
   VAR
      State : Int := 1;
   END_VAR
BEGIN
   CASE #State OF
       1: // Init
           IF #Start THEN
               #State := 2;
           END_IF;
       2:  // Emit pallet
           IF NOT #PalletSensor THEN
               #PalletEmitter := TRUE;
           ELSE
               #PalletEmitter := FALSE;
               #State := 3;
           END_IF;
       3:  // Pallet moving
           #PalletConveyor := #Start;
           #ElevatorConveyor := #Start;
           IF #ElevatorFrontLimit THEN
               #PalletConveyor := FALSE;
               #ElevatorConveyor := FALSE;
               #State := 4;
           END_IF;
       4: // Pallet done;
           IF NOT #ElevatorFrontLimit THEN
               #State := 1;
           END_IF;

   END_CASE;

   #Done := (#State = 4);
END_FUNCTION_BLOCK

FUNCTION_BLOCK "BoxFeedConv"   // FB16, SCL
{ S7_Optimized_Access := 'TRUE' }
VERSION : 0.1
   VAR_INPUT
      EmitSensor : Bool;
      Run : Bool;
      BoxCount : Int;
      StopCount : Int;
      EndSensor : Bool;
      NextBusy : Bool;
   END_VAR
   VAR_OUTPUT
      Conveyor : Bool;
      BoxEmitter : Bool;
   END_VAR
   VAR
      State : Int := 1;
      EmitterSensorNEdge : F_TRIG;
   END_VAR
   VAR_TEMP
      Stop : Bool;
   END_VAR
BEGIN
   #Stop := (#EndSensor AND (#BoxCount = #StopCount)) OR (#NextBusy AND #EndSensor) OR NOT #Run;
   #EmitterSensorNEdge(CLK:=#EmitSensor);
   #BoxEmitter := #EmitSensor;

   CASE #State OF
       1:  //Running
           IF #Stop THEN
               #State := 2;
           END_IF;
       2:  //Stop
           IF NOT #Stop THEN
               #State := 1;
           END_IF;
   END_CASE;

   #Conveyor := (#State = 1);
END_FUNCTION_BLOCK

// folder: StorageCrane

FUNCTION_BLOCK "StorageCrane"   // FB8, SCL
{ S7_Optimized_Access := 'TRUE' }
VERSION : 0.1
   VAR_INPUT
      TargetPosition : Int;
      RequestLoad : Bool;
      RequestUnload : Bool;
      Run : Bool;
   END_VAR
   VAR_OUTPUT
      Busy : Bool;
      LoadDone : Bool;
      UnloadDone : Bool;
   END_VAR
   VAR_IN_OUT
      StorageCraneUDT : "StorageCraneUDT";
   END_VAR
   VAR
      State : Int;
      CraneLoad : "CraneLoad";
      CraneUnload : "CraneUnload";
      LoadIO : "StorageCraneUDT";
      UnloadIO : "StorageCraneUDT";
   END_VAR
BEGIN
   #LoadIO.In := #StorageCraneUDT.In;
   #LoadIO.CraneSides := #StorageCraneUDT.CraneSides;
   #UnloadIO.In := #StorageCraneUDT.In;
   #UnloadIO.CraneSides := #StorageCraneUDT.CraneSides;

   #CraneLoad(TargetPosition := #TargetPosition,
              Start := #RequestLoad AND NOT #RequestUnload AND #Run,
              StorageCraneUDT := #LoadIO);
   #CraneUnload(TargetPosition:=#TargetPosition,
                Start:=#RequestUnload AND NOT #RequestLoad AND #Run,
                StorageCraneUDT:=#UnloadIO); 

   IF #CraneLoad.Busy THEN
       #StorageCraneUDT.Out.Position := #LoadIO.Out.Position;
   ELSIF #CraneUnload.Busy THEN
       #StorageCraneUDT.Out.Position := #UnloadIO.Out.Position;
   END_IF;

   #StorageCraneUDT.Out.Right := #LoadIO.Out.Right OR #UnloadIO.Out.Right;
   #StorageCraneUDT.Out.Left := #LoadIO.Out.Left OR #UnloadIO.Out.Left;
   #StorageCraneUDT.Out.Lift := #LoadIO.Out.Lift OR #UnloadIO.Out.Lift;

   #Busy:=#CraneLoad.Busy OR #CraneUnload.Busy;
   #LoadDone := #CraneLoad.Done;
   #UnloadDone := #CraneUnload.Done;
END_FUNCTION_BLOCK

FUNCTION_BLOCK "CraneLoad"   // FB9, SCL
{ S7_Optimized_Access := 'TRUE' }
VERSION : 0.1
   VAR_INPUT
      TargetPosition : DInt;
      Start : Bool;
   END_VAR
   VAR_OUTPUT
      Busy : Bool;
      Done : Bool;
   END_VAR
   VAR_IN_OUT
      StorageCraneUDT : "StorageCraneUDT";
   END_VAR
   VAR
      State : Int := 1;
      CraneForks : "CraneForks";
      CraneLift : "CraneLift";
      CraneMove : "CraneMove";
   END_VAR
   VAR CONSTANT
      StartPosition : Int := 21474;
   END_VAR
BEGIN
   #CraneForks(LeftLimit:=#StorageCraneUDT.In.LeftLimit,
               MidLimit:=#StorageCraneUDT.In.MidLimit,
               RightLimit:=#StorageCraneUDT.In.RightLimit,
               ExtendLeft=>#StorageCraneUDT.Out.Left,
               ExtendRight=>#StorageCraneUDT.Out.Right);
   #CraneLift(MovingZ:=#StorageCraneUDT.In.MovingZ,
              Lift=>#StorageCraneUDT.Out.Lift);
   #CraneMove(MovingX:=#StorageCraneUDT.In.MovingX,
              MovingZ:=#StorageCraneUDT.In.MovingZ,
              Position=>#StorageCraneUDT.Out.Position);

   CASE #State OF
       1:  // Idle
           #Done := FALSE;
           IF #Start THEN
               #State := 2;
           END_IF;

       2:  // Extend forks to pickup
           #CraneForks.SideRight := #StorageCraneUDT.CraneSides.PickupRight;
           #CraneForks.Extend := TRUE;
           IF #CraneForks.Extended THEN
               #State := 3;
           END_IF;

       3:  // Lift pallet
           #CraneLift.RequestLift := TRUE;
           IF #CraneLift.Done THEN
               #State := 4;
           END_IF;

       4:  // Retract forks
           #CraneForks.Extend := FALSE;
           IF #CraneForks.Retracted THEN
               #State := 5;
           END_IF;

       5:  // Move crane
           #CraneMove.TargetPosition := #TargetPosition;
           #CraneMove.Start := TRUE;
           IF #CraneMove.Done THEN
               #CraneMove.Start := FALSE;
               #State := 6;
           END_IF;

       6:  // Extend forks to load
           #CraneForks.SideRight := #StorageCraneUDT.CraneSides.LoadRight;
           #CraneForks.Extend := TRUE;
           IF #CraneForks.Extended THEN
               #State := 7;
           END_IF;

       7: // Lower pallet
           #CraneLift.RequestLift := FALSE;
           IF #CraneLift.Done THEN
               #State := 8;
           END_IF;

       8:  // Retract forks
           #CraneForks.Extend := FALSE;
           IF #CraneForks.Retracted THEN
               #State := 9;
           END_IF;

       9:  // Back to load zone
           #CraneMove.TargetPosition := #StartPosition;
           #CraneMove.Start := TRUE;
           IF #CraneMove.Done THEN
               #CraneMove.Start := FALSE;
               #State := 1;
               #Done := TRUE;
           END_IF;

   END_CASE;

   #Busy := #State > 1;
END_FUNCTION_BLOCK

FUNCTION_BLOCK "CraneUnload"   // FB10, SCL
{ S7_Optimized_Access := 'TRUE' }
VERSION : 0.1
   VAR_INPUT
      TargetPosition : Int;
      Start : Bool;
   END_VAR
   VAR_OUTPUT
      Busy : Bool;
      Done : Bool;
   END_VAR
   VAR_IN_OUT
      StorageCraneUDT : "StorageCraneUDT";
   END_VAR
   VAR
      State : Int := 1;
      CraneForks : "CraneForks";
      CraneLift : "CraneLift";
      CraneMove : "CraneMove";
   END_VAR
   VAR CONSTANT
      StartPosition : Int := 21474;
   END_VAR
BEGIN
   #CraneForks(LeftLimit:=#StorageCraneUDT.In.LeftLimit,
               MidLimit:=#StorageCraneUDT.In.MidLimit,
               RightLimit:=#StorageCraneUDT.In.RightLimit,
               ExtendLeft=>#StorageCraneUDT.Out.Left,
               ExtendRight=>#StorageCraneUDT.Out.Right);
   #CraneLift(MovingZ:=#StorageCraneUDT.In.MovingZ,
              Lift=>#StorageCraneUDT.Out.Lift);
   #CraneMove(MovingX:=#StorageCraneUDT.In.MovingX,
              MovingZ:=#StorageCraneUDT.In.MovingZ,
              Position=>#StorageCraneUDT.Out.Position);

   CASE #State OF
       1:  // Idle
           #Done := FALSE;
           IF #Start THEN
               #State := 2;
           END_IF;
           ;
       2:  // Move to target position
           #CraneMove.TargetPosition:=#TargetPosition;
           #CraneMove.Start := TRUE;
           IF #CraneMove.Done THEN
               #CraneMove.Start := FALSE;
               #State := 3;
           END_IF;

       3:  // Extend forks
           #CraneForks.Extend := TRUE;
           #CraneForks.SideRight := #StorageCraneUDT.CraneSides.LoadRight;
           IF #CraneForks.Extended THEN
               #State := 4;
           END_IF;

       4:  // Lift pallet
           #CraneLift.RequestLift := TRUE;
           IF #CraneLift.Done THEN
               #State := 5;
           END_IF;

       5:  // Retract forks
           #CraneForks.Extend := FALSE;
           IF #CraneForks.Retracted THEN
               #State := 6;
           END_IF;

       6:  // Move to start position
           #CraneMove.TargetPosition := #StartPosition;
           #CraneMove.Start := TRUE;
           IF #CraneMove.Done THEN
               #CraneMove.Start := FALSE;
               #State := 7;
           END_IF;

       7:  // Extend forks
           #CraneForks.SideRight := #StorageCraneUDT.CraneSides.UnloadRight;
           #CraneForks.Extend := TRUE;
           IF #CraneForks.Extended THEN
               #State := 8;
           END_IF;

       8: // Lower pallet
           #CraneLift.RequestLift := FALSE;
           IF #CraneLift.Done THEN
               #State := 9;
           END_IF;

       9:  // Retract forks
           #CraneForks.Extend := FALSE;
           IF #CraneForks.Retracted THEN
               #State := 1;
               #Done := TRUE;
           END_IF;

   END_CASE;

   #Busy := #State > 1;
END_FUNCTION_BLOCK

FUNCTION_BLOCK "CraneForks"   // FB11, SCL
{ S7_Optimized_Access := 'TRUE' }
VERSION : 0.1
   VAR_INPUT
      LeftLimit : Bool;
      MidLimit : Bool;
      RightLimit : Bool;
      Extend : Bool;
      SideRight : Bool;
   END_VAR
   VAR_OUTPUT
      ExtendLeft : Bool;
      ExtendRight : Bool;
      Retracted : Bool;
      Extended : Bool;
   END_VAR
   VAR
      State : Int;
      SideRightLatched : Bool;
      OppositeRetracted : Bool;
      ActiveExtended : Bool;
   END_VAR
BEGIN
   IF #Extend AND #MidLimit THEN
       #SideRightLatched := #SideRight;
   END_IF;

   IF #SideRightLatched THEN
       #Extended := #Extend AND #RightLimit;
   ELSE
       #Extended := #Extend AND #LeftLimit;
   END_IF;

   #Retracted := (NOT #Extend) AND #MidLimit;
   #ExtendLeft := #Extend AND (NOT #SideRightLatched);
   #ExtendRight := #Extend AND (#SideRightLatched);
END_FUNCTION_BLOCK

FUNCTION_BLOCK "CraneLift"   // FB12, SCL
{ S7_Optimized_Access := 'TRUE' }
VERSION : 0.1
   VAR_INPUT
      RequestLift : Bool;
      MovingZ : Bool;
   END_VAR
   VAR_OUTPUT
      Done : Bool;
      Lift : Bool;
   END_VAR
   VAR
      RequestLiftPEdge : R_TRIG;
      State : Int := 1;
      RequestLiftNEdge : F_TRIG;
   END_VAR
BEGIN
   #Done := FALSE;
   #RequestLiftPEdge(CLK:=#RequestLift);
   #RequestLiftNEdge(CLK:=#RequestLift);

   CASE #State OF
       1:  // Idle
           IF #RequestLiftPEdge.Q THEN
               #Lift := TRUE;
               #State := 2;
           ELSIF #RequestLiftNEdge.Q THEN
               #Lift := FALSE;
               #State := 2;
           END_IF;
           ;
       2:  // WaitStart
           IF #MovingZ THEN
               #State := 3;
           END_IF;
           ;
       3: // Moving
           IF NOT #MovingZ THEN
               #Done := TRUE;
               #State := 1;
           END_IF;
           ;
   END_CASE;
END_FUNCTION_BLOCK

FUNCTION_BLOCK "CraneMove"   // FB13, SCL
{ S7_Optimized_Access := 'TRUE' }
VERSION : 0.1
   VAR_INPUT
      MovingX : Bool;
      MovingZ : Bool;
      Start : Bool;
      TargetPosition : Int;
   END_VAR
   VAR_OUTPUT
      Position : Int := 21474;
      Done : Bool;
   END_VAR
   VAR
      Moving : Bool;
      State : Int := 1;
      StartPEdge : R_TRIG;
   END_VAR
BEGIN
   #Done := FALSE;
   #StartPEdge(CLK:=#Start);
   #Moving := #MovingX OR #MovingZ;

   CASE #State OF
       1:  // Idle
           IF #StartPEdge.Q THEN
               #Position:=#TargetPosition;
               #State := 2;
           END_IF;

       2:  // WaitStart
           IF #Moving THEN
               #State := 3;
           END_IF;

       3: // Moving
           IF NOT #Moving THEN
               #Done := TRUE;
               #State := 1;
           END_IF;

   END_CASE;
END_FUNCTION_BLOCK

// folder: WarehouseManager

FUNCTION_BLOCK "WarehouseManager"   // FB14, SCL
{ S7_Optimized_Access := 'TRUE' }
VERSION : 0.1
   VAR_INPUT
      LoadDone : Array[1..2] of Bool;
      UnloadDone : Array[1..2] of Bool;
      CraneBusy : Array[1..2] of Bool;
      PalletReady : Bool;
      UnloadRequest : Bool;
      UnloadRack : Int;
      UnloadSlot : Int;
      Run : Bool;
   END_VAR
   VAR_OUTPUT
      Full : Bool;
      Busy : Bool;
      PalletStored : Bool;
      PalletUnloaded : Bool;
      UnloadRejected : Bool;
      LoadStart : Array[1..2] of Bool;
      UnloadStart : Array[1..2] of Bool;
      TargetSlot : Array[1..2] of Int;
      Rack : Int;
      CraneStatus : Array[1..2] of Int;
   END_VAR
   VAR_IN_OUT
      Rack1Slots : Array[*] of "WarehouseSlotUDT";
      Rack2Slots : Array[*] of "WarehouseSlotUDT";
   END_VAR
   VAR
      LoadManager : "LoadManager";
      UnloadManager : "UnloadManager";
   END_VAR
   VAR_TEMP
      i : Int;
      loadFree : Array[1..2] of Bool;
      unloadFree : Array[1..2] of Bool;
   END_VAR
BEGIN
   FOR #i := 1 TO 2 DO
       #loadFree[#i] := (NOT #CraneBusy[#i]) AND (NOT #UnloadManager.Active[#i]);
   END_FOR;

   #LoadManager(PalletReady:=#PalletReady,
                LoadDone:=#LoadDone,
                CraneFree:=#loadFree,
                Run:=#Run,
                Rack=>#Rack,
                Rack1Slots:=#Rack1Slots,
                Rack2Slots:=#Rack2Slots); 

   FOR #i := 1 TO 2 DO
       #unloadFree[#i] := (NOT #CraneBusy[#i]) AND (NOT #LoadManager.Active[#i]);
   END_FOR;

   #UnloadManager(UnloadRequest:=#UnloadRequest,
                  Run:=#Run,
                  UnloadRack:=#UnloadRack,
                  UnloadSlot:=#UnloadSlot,
                  UnloadDone:=#UnloadDone,
                  CraneFree:=#unloadFree,
                  Rack1Slots:=#Rack1Slots,
                  Rack2Slots:=#Rack2Slots);

   FOR #i := 1 TO 2 DO
       #LoadStart[#i] := #LoadManager.LoadStart[#i];
       #UnloadStart[#i] := #UnloadManager.UnloadStart[#i];

       IF #UnloadManager.Active[#i] THEN
           #TargetSlot[#i] := #UnloadManager.TargetSlot[#i];
       ELSE
           #TargetSlot[#i] := #LoadManager.TargetSlot[#i];
       END_IF;
   END_FOR;

   FOR #i := 1 TO 2 DO
       IF NOT #CraneBusy[#i] THEN
           #CraneStatus[#i] := 0;
       ELSIF #CraneBusy[#i] AND #LoadManager.Active[#i] AND (NOT #UnloadManager.Active[#i]) THEN
           #CraneStatus[#i] := 1;
       ELSIF #CraneBusy[#i] AND #UnloadManager.Active[#i] AND (NOT #UnloadManager.Active[#i]) THEN
           #CraneStatus[#i] := 2;
       END_IF;
   END_FOR;

   #Busy := #LoadManager.Busy OR #UnloadManager.Busy;
   #Full := #LoadManager.Full;
   #UnloadRejected := #UnloadManager.UnloadRejected;
END_FUNCTION_BLOCK

FUNCTION_BLOCK "LoadManager"   // FB17, SCL
{ S7_Optimized_Access := 'TRUE' }
VERSION : 0.1
   VAR_INPUT
      PalletReady : Bool;
      LoadDone : Array[1..2] of Bool;
      CraneFree : Array[1..2] of Bool;
      Run : Bool;
   END_VAR
   VAR_OUTPUT
      Busy : Bool;
      Full : Bool;
      PalletStored : Bool;
      Rack : Int;
      LoadStart : Array[1..2] of Bool;
      Active : Array[1..2] of Bool;
      TargetSlot : Array[1..2] of Int;
   END_VAR
   VAR_IN_OUT
      Rack1Slots : Array[*] of "WarehouseSlotUDT";
      Rack2Slots : Array[*] of "WarehouseSlotUDT";
   END_VAR
   VAR
      State : Int := 1;
      NextPalletId : Int;
      CurrentId : Int;
      Slot : Int;
      LastRack : Int;
      PalletPending : Bool;
      CpuTime : DTL;
      PalletReadyPEdge : R_TRIG;
   END_VAR
   VAR_TEMP
      temptime : Int;
      realfree1 : Int;
      realfree2 : Int;
      free1 : Int;
      free2 : Int;
      i : Int;
   END_VAR
BEGIN
   #PalletReadyPEdge(CLK:=#PalletReady);
   #temptime := RD_LOC_T(OUT => #CpuTime);
   IF #PalletReadyPEdge.Q THEN
       #PalletPending := TRUE;
   END_IF;

   CASE #State OF

       1: // Idle
           IF #PalletPending AND #Run THEN
               #realfree1 := "CountFreeSlots"(Slots := #Rack1Slots);
               #realfree2 := "CountFreeSlots"(Slots := #Rack2Slots);

               IF #CraneFree[1] THEN
                   #free1 := #realfree1;
               ELSE
                   #free1 := 0;
               END_IF;

               IF #CraneFree[2] THEN
                   #free2 := #realfree2;
               ELSE
                   #free2 := 0;
               END_IF;

               #Rack := "SelectRack"(FreeSlotsRack1 := #realfree1, FreeSlotsRack2 := #realfree2, Last := #LastRack);

               IF #Rack = 0 THEN
                   #Full := (#realfree1 = 0) AND (#realfree2 = 0);
               ELSE
                   #PalletPending := FALSE;
                   #NextPalletId := #NextPalletId + 1;
                   #CurrentId := #NextPalletId;
                   IF #Rack = 1 THEN
                       #Slot := "ReserveFirstFree"(Slot := #Rack1Slots, PalletId := #CurrentId);
                   ELSIF #Rack = 2 THEN
                       #Slot := "ReserveFirstFree"(Slot := #Rack2Slots, PalletId := #CurrentId);
                   END_IF;
                   #State := 2;
               END_IF;
           END_IF;

       2:  // Loading
           #LoadStart[#Rack] := TRUE;
           #TargetSlot[#Rack] := #Slot;

           IF #LoadDone[#Rack] THEN
               IF #Rack = 1 THEN
                   #Rack1Slots[#Slot].Status := 2;
                   #Rack1Slots[#Slot]."Time" := #CpuTime;
               ELSIF #Rack = 2 THEN
                   #Rack2Slots[#Slot].Status := 2;
                   #Rack2Slots[#Slot]."Time" := #CpuTime;
               END_IF;
               #PalletStored := TRUE;
               #LoadStart[#Rack] := FALSE;
               #State := 1;
           END_IF;

   END_CASE;

   FOR #i := 1 TO 2 DO
       #Active[#i] := (#State = 2) AND (#Rack = #i);
   END_FOR;

   #Busy := #State = 2 OR #PalletPending;
END_FUNCTION_BLOCK

FUNCTION_BLOCK "UnloadManager"   // FB18, SCL
{ S7_Optimized_Access := 'TRUE' }
VERSION : 0.1
   VAR_INPUT
      UnloadRequest : Bool;
      Run : Bool;
      UnloadRack : Int;
      UnloadSlot : Int;
      UnloadDone : Array[1..2] of Bool;
      CraneFree : Array[1..2] of Bool;
   END_VAR
   VAR_OUTPUT
      UnloadStart : Array[1..2] of Bool;
      Active : Array[1..2] of Bool;
      TargetSlot : Array[1..2] of Int;
      Busy : Bool;
      PalletUnloaded : Bool;
      UnloadRejected : Bool;
   END_VAR
   VAR_IN_OUT
      Rack1Slots : Array[*] of "WarehouseSlotUDT";
      Rack2Slots : Array[*] of "WarehouseSlotUDT";
   END_VAR
   VAR
      State : Int := 1;
      UnloadId : Int;
      Rack : Int;
      Slot : Int;
      UnloadPending : Bool;
      RequestedRack : Int;
      RequestedSlot : Int;
      UnloadRequestPEdge : R_TRIG;
   END_VAR
   VAR_TEMP
      i : Int;
      id : Int;
   END_VAR
BEGIN
   #UnloadRequestPEdge(CLK:=#UnloadRequest);

   IF #UnloadRequestPEdge.Q THEN
       #UnloadPending := TRUE;
       #RequestedRack := #UnloadRack;
       #RequestedSlot := #UnloadSlot;
   END_IF;

   CASE #State OF
       1: // Idle
           IF #UnloadPending AND #Run THEN
               IF #CraneFree[#RequestedRack] THEN
                   #UnloadPending := FALSE;
                   #id := 0;
                   IF #RequestedRack = 1 THEN
                       #id := "ReserveUnload"(Slot := #RequestedSlot, Slots := #Rack1Slots);
                   ELSIF #RequestedRack = 2 THEN
                       #id := "ReserveUnload"(Slot := #RequestedSlot, Slots := #Rack2Slots);
                   END_IF;

                   IF #id > 0 THEN
                       #Rack := #RequestedRack;
                       #Slot := #RequestedSlot;
                       #UnloadId := #id;
                       #State := 2;
                   ELSE
                       #UnloadRejected := TRUE;
                   END_IF;
               END_IF;
           END_IF;

       2: // Unloading
           #UnloadStart[#Rack] := TRUE;
           #TargetSlot[#Rack] := #Slot;

           IF #UnloadDone[#Rack] THEN
               IF #Rack = 1 THEN
                   #Rack1Slots[#Slot].Status := 0;
                   #Rack1Slots[#Slot].Id := 0;
                   #Rack1Slots[#Slot]."Time" := DTL#1970-01-01-00:00:00;
               ELSIF #Rack = 2 THEN
                   #Rack2Slots[#Slot].Status := 0;
                   #Rack2Slots[#Slot].Id := 0;
                   #Rack2Slots[#Slot]."Time" := DTL#1970-01-01-00:00:00;
               END_IF;
               #PalletUnloaded := TRUE;
               #UnloadStart[#Rack] := FALSE;
               #State := 1;
           END_IF;

   END_CASE;

   FOR #i := 1 TO 2 DO
       #Active[#i] := (#State = 2) AND (#Rack = #i);
   END_FOR;

   #Busy := #State = 2 OR #UnloadPending;
END_FUNCTION_BLOCK

FUNCTION "CountFreeSlots" : Int   // FC1, SCL
{ S7_Optimized_Access := 'TRUE' }
VERSION : 0.1
   VAR_IN_OUT
      Slots : Array[*] of "WarehouseSlotUDT";
   END_VAR
   VAR_TEMP
      i : Int;
      n : Int;
   END_VAR
BEGIN
   #n := 0;
   FOR #i := 1 TO 54 DO
       IF #Slots[#i].Status=0 THEN
           #n := #n + 1;
       END_IF;
   END_FOR;

   #CountFreeSlots := #n;
END_FUNCTION

FUNCTION "ReserveFirstFree" : Int   // FC2, SCL
{ S7_Optimized_Access := 'TRUE' }
VERSION : 0.1
   VAR_INPUT
      PalletId : Int;
   END_VAR
   VAR_IN_OUT
      Slot : Array[*] of "WarehouseSlotUDT";
   END_VAR
   VAR_TEMP
      i : Int;
   END_VAR
BEGIN
   #ReserveFirstFree := 0;

   FOR #i := 1 TO 54 DO
       IF #Slot[#i].Status = 0 THEN
           #Slot[#i].Status := 1;
           #Slot[#i].Id := #PalletId;
           #ReserveFirstFree := #i;
           EXIT;
       END_IF;
   END_FOR;
END_FUNCTION

FUNCTION "SelectRack" : Int   // FC3, SCL
{ S7_Optimized_Access := 'TRUE' }
VERSION : 0.1
   VAR_INPUT
      FreeSlotsRack1 : Int;
      FreeSlotsRack2 : Int;
   END_VAR
   VAR_IN_OUT
      Last : Int;
   END_VAR
BEGIN
   IF (#FreeSlotsRack1 > 0) AND (#FreeSlotsRack2 > 0) THEN
       IF #FreeSlotsRack1 > #FreeSlotsRack2 THEN
           #SelectRack := 1;
       ELSIF #FreeSlotsRack2 > #FreeSlotsRack1 THEN
           #SelectRack := 2;
       ELSIF #Last = 1 THEN
           #SelectRack := 2;
       ELSE
           #SelectRack := 1;
       END_IF;
   ELSIF #FreeSlotsRack1 > 0 THEN
       #SelectRack := 1;
   ELSIF #FreeSlotsRack2 > 0 THEN
       #SelectRack := 2;
   ELSE
       #SelectRack := 0;
   END_IF;

   IF #SelectRack <> 0 THEN
       #Last := #SelectRack;
   END_IF;
END_FUNCTION

FUNCTION "ReserveUnload" : Int   // FC7, SCL
{ S7_Optimized_Access := 'TRUE' }
VERSION : 0.1
   VAR_INPUT
      Slot : Int;
   END_VAR
   VAR_IN_OUT
      Slots : Array[*] of "WarehouseSlotUDT";
   END_VAR
BEGIN
   #ReserveUnload := 0;

   IF #Slots[#Slot].Status = 2 THEN
       #Slots[#Slot].Status := 1;
       #ReserveUnload := #Slots[#Slot].Id;
   END_IF;
END_FUNCTION

(* ===== HMI "HMI_RT_1" =====
system functions are stored by id; their names below are inferred from use
connection "HMI_Connection_1": ETHERNET, S7_1500_OMS

HMI tags "Default tag table"
   "WarehouseData_Rack1{1}" : WarehouseSlotUDT = PLC WarehouseData.Rack1[1], 1 s
   "WarehouseData_Rack1{2}" : WarehouseSlotUDT = PLC WarehouseData.Rack1[2], 1 s
   "WarehouseData_Rack1{3}" : WarehouseSlotUDT = PLC WarehouseData.Rack1[3], 1 s
   "WarehouseData_Rack1{4}" : WarehouseSlotUDT = PLC WarehouseData.Rack1[4], 1 s
   "WarehouseData_Rack1{5}" : WarehouseSlotUDT = PLC WarehouseData.Rack1[5], 1 s
   "WarehouseData_Rack1{6}" : WarehouseSlotUDT = PLC WarehouseData.Rack1[6], 1 s
   "WarehouseData_Rack1{7}" : WarehouseSlotUDT = PLC WarehouseData.Rack1[7], 1 s
   "WarehouseData_Rack1{8}" : WarehouseSlotUDT = PLC WarehouseData.Rack1[8], 1 s
   "WarehouseData_Rack1{9}" : WarehouseSlotUDT = PLC WarehouseData.Rack1[9], 1 s
   "WarehouseData_Rack1{10}" : WarehouseSlotUDT = PLC WarehouseData.Rack1[10], 1 s
   "WarehouseData_Rack1{11}" : WarehouseSlotUDT = PLC WarehouseData.Rack1[11], 1 s
   "WarehouseData_Rack1{12}" : WarehouseSlotUDT = PLC WarehouseData.Rack1[12], 1 s
   "WarehouseData_Rack1{13}" : WarehouseSlotUDT = PLC WarehouseData.Rack1[13], 1 s
   "WarehouseData_Rack1{14}" : WarehouseSlotUDT = PLC WarehouseData.Rack1[14], 1 s
   "WarehouseData_Rack1{15}" : WarehouseSlotUDT = PLC WarehouseData.Rack1[15], 1 s
   "WarehouseData_Rack1{16}" : WarehouseSlotUDT = PLC WarehouseData.Rack1[16], 1 s
   "WarehouseData_Rack1{17}" : WarehouseSlotUDT = PLC WarehouseData.Rack1[17], 1 s
   "WarehouseData_Rack1{18}" : WarehouseSlotUDT = PLC WarehouseData.Rack1[18], 1 s
   "WarehouseData_Rack1{19}" : WarehouseSlotUDT = PLC WarehouseData.Rack1[19], 1 s
   "WarehouseData_Rack1{20}" : WarehouseSlotUDT = PLC WarehouseData.Rack1[20], 1 s
   "WarehouseData_Rack1{21}" : WarehouseSlotUDT = PLC WarehouseData.Rack1[21], 1 s
   "WarehouseData_Rack1{22}" : WarehouseSlotUDT = PLC WarehouseData.Rack1[22], 1 s
   "WarehouseData_Rack1{23}" : WarehouseSlotUDT = PLC WarehouseData.Rack1[23], 1 s
   "WarehouseData_Rack1{24}" : WarehouseSlotUDT = PLC WarehouseData.Rack1[24], 1 s
   "WarehouseData_Rack1{25}" : WarehouseSlotUDT = PLC WarehouseData.Rack1[25], 1 s
   "WarehouseData_Rack1{26}" : WarehouseSlotUDT = PLC WarehouseData.Rack1[26], 1 s
   "WarehouseData_Rack1{27}" : WarehouseSlotUDT = PLC WarehouseData.Rack1[27], 1 s
   "WarehouseData_Rack1{28}" : WarehouseSlotUDT = PLC WarehouseData.Rack1[28], 1 s
   "WarehouseData_Rack1{29}" : WarehouseSlotUDT = PLC WarehouseData.Rack1[29], 1 s
   "WarehouseData_Rack1{30}" : WarehouseSlotUDT = PLC WarehouseData.Rack1[30], 1 s
   "WarehouseData_Rack1{31}" : WarehouseSlotUDT = PLC WarehouseData.Rack1[31], 1 s
   "WarehouseData_Rack1{32}" : WarehouseSlotUDT = PLC WarehouseData.Rack1[32], 1 s
   "WarehouseData_Rack1{33}" : WarehouseSlotUDT = PLC WarehouseData.Rack1[33], 1 s
   "WarehouseData_Rack1{34}" : WarehouseSlotUDT = PLC WarehouseData.Rack1[34], 1 s
   "WarehouseData_Rack1{35}" : WarehouseSlotUDT = PLC WarehouseData.Rack1[35], 1 s
   "WarehouseData_Rack1{36}" : WarehouseSlotUDT = PLC WarehouseData.Rack1[36], 1 s
   "WarehouseData_Rack1{37}" : WarehouseSlotUDT = PLC WarehouseData.Rack1[37], 1 s
   "WarehouseData_Rack1{38}" : WarehouseSlotUDT = PLC WarehouseData.Rack1[38], 1 s
   "WarehouseData_Rack1{39}" : WarehouseSlotUDT = PLC WarehouseData.Rack1[39], 1 s
   "WarehouseData_Rack1{40}" : WarehouseSlotUDT = PLC WarehouseData.Rack1[40], 1 s
   "WarehouseData_Rack1{41}" : WarehouseSlotUDT = PLC WarehouseData.Rack1[41], 1 s
   "WarehouseData_Rack1{42}" : WarehouseSlotUDT = PLC WarehouseData.Rack1[42], 1 s
   "WarehouseData_Rack1{43}" : WarehouseSlotUDT = PLC WarehouseData.Rack1[43], 1 s
   "WarehouseData_Rack1{44}" : WarehouseSlotUDT = PLC WarehouseData.Rack1[44], 1 s
   "WarehouseData_Rack1{45}" : WarehouseSlotUDT = PLC WarehouseData.Rack1[45], 1 s
   "WarehouseData_Rack1{46}" : WarehouseSlotUDT = PLC WarehouseData.Rack1[46], 1 s
   "WarehouseData_Rack1{47}" : WarehouseSlotUDT = PLC WarehouseData.Rack1[47], 1 s
   "WarehouseData_Rack1{48}" : WarehouseSlotUDT = PLC WarehouseData.Rack1[48], 1 s
   "WarehouseData_Rack1{49}" : WarehouseSlotUDT = PLC WarehouseData.Rack1[49], 1 s
   "WarehouseData_Rack1{50}" : WarehouseSlotUDT = PLC WarehouseData.Rack1[50], 1 s
   "WarehouseData_Rack1{51}" : WarehouseSlotUDT = PLC WarehouseData.Rack1[51], 1 s
   "WarehouseData_Rack1{52}" : WarehouseSlotUDT = PLC WarehouseData.Rack1[52], 1 s
   "WarehouseData_Rack1{53}" : WarehouseSlotUDT = PLC WarehouseData.Rack1[53], 1 s
   "WarehouseData_Rack1{54}" : WarehouseSlotUDT = PLC WarehouseData.Rack1[54], 1 s
   "WarehouseData_Rack2{1}" : WarehouseSlotUDT = PLC WarehouseData.Rack2[1] AT %DB1.DBW0, 1 s
   "WarehouseData_Rack2{2}" : WarehouseSlotUDT = PLC WarehouseData.Rack2[2] AT %DB1.DBW0, 1 s
   "WarehouseData_Rack2{3}" : WarehouseSlotUDT = PLC WarehouseData.Rack2[3] AT %DB1.DBW0, 1 s
   "WarehouseData_Rack2{4}" : WarehouseSlotUDT = PLC WarehouseData.Rack2[4] AT %DB1.DBW0, 1 s
   "WarehouseData_Rack2{5}" : WarehouseSlotUDT = PLC WarehouseData.Rack2[5] AT %DB1.DBW0, 1 s
   "WarehouseData_Rack2{6}" : WarehouseSlotUDT = PLC WarehouseData.Rack2[6] AT %DB1.DBW0, 1 s
   "WarehouseData_Rack2{7}" : WarehouseSlotUDT = PLC WarehouseData.Rack2[7] AT %DB1.DBW0, 1 s
   "WarehouseData_Rack2{8}" : WarehouseSlotUDT = PLC WarehouseData.Rack2[8] AT %DB1.DBW0, 1 s
   "WarehouseData_Rack2{9}" : WarehouseSlotUDT = PLC WarehouseData.Rack2[9] AT %DB1.DBW0, 1 s
   "WarehouseData_Rack2{10}" : WarehouseSlotUDT = PLC WarehouseData.Rack2[10] AT %DB1.DBW0, 1 s
   "WarehouseData_Rack2{11}" : WarehouseSlotUDT = PLC WarehouseData.Rack2[11] AT %DB1.DBW0, 1 s
   "WarehouseData_Rack2{12}" : WarehouseSlotUDT = PLC WarehouseData.Rack2[12] AT %DB1.DBW0, 1 s
   "WarehouseData_Rack2{13}" : WarehouseSlotUDT = PLC WarehouseData.Rack2[13] AT %DB1.DBW0, 1 s
   "WarehouseData_Rack2{14}" : WarehouseSlotUDT = PLC WarehouseData.Rack2[14] AT %DB1.DBW0, 1 s
   "WarehouseData_Rack2{15}" : WarehouseSlotUDT = PLC WarehouseData.Rack2[15] AT %DB1.DBW0, 1 s
   "WarehouseData_Rack2{16}" : WarehouseSlotUDT = PLC WarehouseData.Rack2[16] AT %DB1.DBW0, 1 s
   "WarehouseData_Rack2{17}" : WarehouseSlotUDT = PLC WarehouseData.Rack2[17] AT %DB1.DBW0, 1 s
   "WarehouseData_Rack2{18}" : WarehouseSlotUDT = PLC WarehouseData.Rack2[18] AT %DB1.DBW0, 1 s
   "WarehouseData_Rack2{19}" : WarehouseSlotUDT = PLC WarehouseData.Rack2[19] AT %DB1.DBW0, 1 s
   "WarehouseData_Rack2{20}" : WarehouseSlotUDT = PLC WarehouseData.Rack2[20] AT %DB1.DBW0, 1 s
   "WarehouseData_Rack2{21}" : WarehouseSlotUDT = PLC WarehouseData.Rack2[21] AT %DB1.DBW0, 1 s
   "WarehouseData_Rack2{22}" : WarehouseSlotUDT = PLC WarehouseData.Rack2[22] AT %DB1.DBW0, 1 s
   "WarehouseData_Rack2{23}" : WarehouseSlotUDT = PLC WarehouseData.Rack2[23] AT %DB1.DBW0, 1 s
   "WarehouseData_Rack2{24}" : WarehouseSlotUDT = PLC WarehouseData.Rack2[24] AT %DB1.DBW0, 1 s
   "WarehouseData_Rack2{25}" : WarehouseSlotUDT = PLC WarehouseData.Rack2[25] AT %DB1.DBW0, 1 s
   "WarehouseData_Rack2{26}" : WarehouseSlotUDT = PLC WarehouseData.Rack2[26] AT %DB1.DBW0, 1 s
   "WarehouseData_Rack2{27}" : WarehouseSlotUDT = PLC WarehouseData.Rack2[27] AT %DB1.DBW0, 1 s
   "WarehouseData_Rack2{28}" : WarehouseSlotUDT = PLC WarehouseData.Rack2[28] AT %DB1.DBW0, 1 s
   "WarehouseData_Rack2{29}" : WarehouseSlotUDT = PLC WarehouseData.Rack2[29] AT %DB1.DBW0, 1 s
   "WarehouseData_Rack2{30}" : WarehouseSlotUDT = PLC WarehouseData.Rack2[30] AT %DB1.DBW0, 1 s
   "WarehouseData_Rack2{31}" : WarehouseSlotUDT = PLC WarehouseData.Rack2[31] AT %DB1.DBW0, 1 s
   "WarehouseData_Rack2{32}" : WarehouseSlotUDT = PLC WarehouseData.Rack2[32] AT %DB1.DBW0, 1 s
   "WarehouseData_Rack2{33}" : WarehouseSlotUDT = PLC WarehouseData.Rack2[33] AT %DB1.DBW0, 1 s
   "WarehouseData_Rack2{34}" : WarehouseSlotUDT = PLC WarehouseData.Rack2[34] AT %DB1.DBW0, 1 s
   "WarehouseData_Rack2{35}" : WarehouseSlotUDT = PLC WarehouseData.Rack2[35] AT %DB1.DBW0, 1 s
   "WarehouseData_Rack2{36}" : WarehouseSlotUDT = PLC WarehouseData.Rack2[36] AT %DB1.DBW0, 1 s
   "WarehouseData_Rack2{37}" : WarehouseSlotUDT = PLC WarehouseData.Rack2[37] AT %DB1.DBW0, 1 s
   "WarehouseData_Rack2{38}" : WarehouseSlotUDT = PLC WarehouseData.Rack2[38] AT %DB1.DBW0, 1 s
   "WarehouseData_Rack2{39}" : WarehouseSlotUDT = PLC WarehouseData.Rack2[39] AT %DB1.DBW0, 1 s
   "WarehouseData_Rack2{40}" : WarehouseSlotUDT = PLC WarehouseData.Rack2[40] AT %DB1.DBW0, 1 s
   "WarehouseData_Rack2{41}" : WarehouseSlotUDT = PLC WarehouseData.Rack2[41] AT %DB1.DBW0, 1 s
   "WarehouseData_Rack2{42}" : WarehouseSlotUDT = PLC WarehouseData.Rack2[42] AT %DB1.DBW0, 1 s
   "WarehouseData_Rack2{43}" : WarehouseSlotUDT = PLC WarehouseData.Rack2[43] AT %DB1.DBW0, 1 s
   "WarehouseData_Rack2{44}" : WarehouseSlotUDT = PLC WarehouseData.Rack2[44] AT %DB1.DBW0, 1 s
   "WarehouseData_Rack2{45}" : WarehouseSlotUDT = PLC WarehouseData.Rack2[45] AT %DB1.DBW0, 1 s
   "WarehouseData_Rack2{46}" : WarehouseSlotUDT = PLC WarehouseData.Rack2[46] AT %DB1.DBW0, 1 s
   "WarehouseData_Rack2{47}" : WarehouseSlotUDT = PLC WarehouseData.Rack2[47] AT %DB1.DBW0, 1 s
   "WarehouseData_Rack2{48}" : WarehouseSlotUDT = PLC WarehouseData.Rack2[48] AT %DB1.DBW0, 1 s
   "WarehouseData_Rack2{49}" : WarehouseSlotUDT = PLC WarehouseData.Rack2[49] AT %DB1.DBW0, 1 s
   "WarehouseData_Rack2{50}" : WarehouseSlotUDT = PLC WarehouseData.Rack2[50] AT %DB1.DBW0, 1 s
   "WarehouseData_Rack2{51}" : WarehouseSlotUDT = PLC WarehouseData.Rack2[51] AT %DB1.DBW0, 1 s
   "WarehouseData_Rack2{52}" : WarehouseSlotUDT = PLC WarehouseData.Rack2[52] AT %DB1.DBW0, 1 s
   "WarehouseData_Rack2{53}" : WarehouseSlotUDT = PLC WarehouseData.Rack2[53] AT %DB1.DBW0, 1 s
   "WarehouseData_Rack2{54}" : WarehouseSlotUDT = PLC WarehouseData.Rack2[54] AT %DB1.DBW0, 1 s
   "SelectedRack" : Int = PLC HMI_Data.SelectedRack AT %DB1.DBW0, 1 s
   "SelectedSlot" : Int = PLC HMI_Data.SelectedSlot AT %DB1.DBW0, 1 s
   "TargetSlot" : WarehouseSlotUDT = PLC HMI_Data.TargetSlot AT %DB1.DBW0, 1 s
   "RetrievePallet" : Bool = PLC HMI_Data.RetrievePallet AT %DB1.DBX0.0, 1 s
   "RacksFull" : Bool = PLC HMI_Data.RacksFull, 1 s
   "CraneStatus" : Array [0..1] of Int = PLC HMI_Data.CraneStatus, 1 s
   "OccupiedSlots" : Array [0..1] of Int = PLC HMI_Data.OccupiedSlots, 1 s
   "StartCmd" : Bool = PLC HMI_Data.StartCmd AT %DB1.DBX0.0, 1 s
   "StopCmd" : Bool = PLC HMI_Data.StopCmd AT %DB1.DBX0.0, 1 s

text list "CraneStatus": 0 'Idle'; 1 'Loading...'; 2 'Unloading...'

text list "SlotStatus": 0 'Empty'; 1 'Reserved'; 2 'Occupied'

screen "Rack 1" 640x480
   Button "Button_1" at 0,0 size 90x66; TextOff 'Rack 1'
      on Click: ActivateScreen("Rack 1", 0)
   Button "Button_2" at 130,0 size 90x66; TextOff 'Rack 2'
      on Click: ActivateScreen("Rack 2", 0)
   DateTimeField "Date/time field_1" at 444,15 size 177x31
   TextField "Text field_46" at 350,88 size 74x28; Text 'Rack 1'
   ScreenModuleView "RackSlot_1" at 562,360 size 44x36; Guid_{11997190-21654} '0'; ScreenModuleType ""
      Guid_{11997190-21133} <- "WarehouseData_Rack1{1}"
      on Guid_{11997190-21491}: function_efd93a16("RackSlotData", 0, 0, -1, -1, 1)
   ScreenModuleView "RackSlot_2" at 512,360 size 44x36; Guid_{11997190-21654} '0'; ScreenModuleType ""
      on Guid_{11997190-21491}: function_efd93a16("RackSlotData", 0, 0, -1, -1, 1)
      Guid_{11997190-21133} <- "WarehouseData_Rack1{1}"
   ScreenModuleView "RackSlot_3" at 562,360 size 44x36; Guid_{11997190-21654} '1'; Guid_{11997190-23841} '1'; ScreenModuleType ""
      on Guid_{11997190-21491}: SetTag("SelectedRack", 1); SetTag("SelectedSlot", 1); function_efd93a16("RackSlotData", 220, 150, -1, -1, 1)
      Guid_{11997190-21133} <- "WarehouseData_Rack1{1}"
   ScreenModuleView "RackSlot_4" at 512,360 size 44x36; Guid_{11997190-21654} '2'; Guid_{11997190-23841} '2'; ScreenModuleType ""
      on Guid_{11997190-21491}: SetTag("SelectedRack", 1); SetTag("SelectedSlot", 2); function_efd93a16("RackSlotData", 220, 150, -1, -1, 1)
      Guid_{11997190-21133} <- "WarehouseData_Rack1{2}"
   ScreenModuleView "RackSlot_5" at 462,360 size 44x36; Guid_{11997190-21654} '3'; Guid_{11997190-23841} '3'; ScreenModuleType ""
      on Guid_{11997190-21491}: SetTag("SelectedRack", 1); SetTag("SelectedSlot", 3); function_efd93a16("RackSlotData", 220, 150, -1, -1, 1)
      Guid_{11997190-21133} <- "WarehouseData_Rack1{3}"
   ScreenModuleView "RackSlot_6" at 412,360 size 44x36; Guid_{11997190-21654} '4'; Guid_{11997190-23841} '4'; ScreenModuleType ""
      on Guid_{11997190-21491}: SetTag("SelectedRack", 1); SetTag("SelectedSlot", 4); function_efd93a16("RackSlotData", 220, 150, -1, -1, 1)
      Guid_{11997190-21133} <- "WarehouseData_Rack1{4}"
   ScreenModuleView "RackSlot_7" at 362,360 size 44x36; Guid_{11997190-21654} '5'; Guid_{11997190-23841} '5'; ScreenModuleType ""
      on Guid_{11997190-21491}: SetTag("SelectedRack", 1); SetTag("SelectedSlot", 5); function_efd93a16("RackSlotData", 220, 150, -1, -1, 1)
      Guid_{11997190-21133} <- "WarehouseData_Rack1{5}"
   ScreenModuleView "RackSlot_8" at 312,360 size 44x36; Guid_{11997190-21654} '6'; Guid_{11997190-23841} '6'; ScreenModuleType ""
      on Guid_{11997190-21491}: SetTag("SelectedRack", 1); SetTag("SelectedSlot", 6); function_efd93a16("RackSlotData", 220, 150, -1, -1, 1)
      Guid_{11997190-21133} <- "WarehouseData_Rack1{6}"
   ScreenModuleView "RackSlot_9" at 262,360 size 44x36; Guid_{11997190-21654} '7'; Guid_{11997190-23841} '7'; ScreenModuleType ""
      on Guid_{11997190-21491}: SetTag("SelectedRack", 1); SetTag("SelectedSlot", 7); function_efd93a16("RackSlotData", 220, 150, -1, -1, 1)
      Guid_{11997190-21133} <- "WarehouseData_Rack1{7}"
   ScreenModuleView "RackSlot_10" at 212,360 size 44x36; Guid_{11997190-21654} '8'; Guid_{11997190-23841} '8'; ScreenModuleType ""
      on Guid_{11997190-21491}: SetTag("SelectedRack", 1); SetTag("SelectedSlot", 8); function_efd93a16("RackSlotData", 220, 150, -1, -1, 1)
      Guid_{11997190-21133} <- "WarehouseData_Rack1{8}"
   ScreenModuleView "RackSlot_11" at 162,360 size 44x36; Guid_{11997190-21654} '9'; Guid_{11997190-23841} '9'; ScreenModuleType ""
      on Guid_{11997190-21491}: SetTag("SelectedRack", 1); SetTag("SelectedSlot", 9); function_efd93a16("RackSlotData", 220, 150, -1, -1, 1)
      Guid_{11997190-21133} <- "WarehouseData_Rack1{9}"
   ScreenModuleView "RackSlot_12" at 562,315 size 44x36; Guid_{11997190-21654} '10'; Guid_{11997190-23841} '10'; ScreenModuleType ""
      on Guid_{11997190-21491}: SetTag("SelectedRack", 1); SetTag("SelectedSlot", 10); function_efd93a16("RackSlotData", 220, 150, -1, -1, 1)
      Guid_{11997190-21133} <- "WarehouseData_Rack1{10}"
   ScreenModuleView "RackSlot_13" at 512,315 size 44x36; Guid_{11997190-21654} '11'; Guid_{11997190-23841} '11'; ScreenModuleType ""
      on Guid_{11997190-21491}: SetTag("SelectedRack", 1); SetTag("SelectedSlot", 11); function_efd93a16("RackSlotData", 220, 150, -1, -1, 1)
      Guid_{11997190-21133} <- "WarehouseData_Rack1{11}"
   ScreenModuleView "RackSlot_14" at 462,315 size 44x36; Guid_{11997190-21654} '12'; Guid_{11997190-23841} '12'; ScreenModuleType ""
      on Guid_{11997190-21491}: SetTag("SelectedRack", 1); SetTag("SelectedSlot", 12); function_efd93a16("RackSlotData", 220, 150, -1, -1, 1)
      Guid_{11997190-21133} <- "WarehouseData_Rack1{12}"
   ScreenModuleView "RackSlot_15" at 412,315 size 44x36; Guid_{11997190-21654} '13'; Guid_{11997190-23841} '13'; ScreenModuleType ""
      on Guid_{11997190-21491}: SetTag("SelectedRack", 1); SetTag("SelectedSlot", 13); function_efd93a16("RackSlotData", 220, 150, -1, -1, 1)
      Guid_{11997190-21133} <- "WarehouseData_Rack1{13}"
   ScreenModuleView "RackSlot_16" at 362,315 size 44x36; Guid_{11997190-21654} '14'; Guid_{11997190-23841} '14'; ScreenModuleType ""
      on Guid_{11997190-21491}: SetTag("SelectedRack", 1); SetTag("SelectedSlot", 14); function_efd93a16("RackSlotData", 220, 150, -1, -1, 1)
      Guid_{11997190-21133} <- "WarehouseData_Rack1{14}"
   ScreenModuleView "RackSlot_17" at 312,315 size 44x36; Guid_{11997190-21654} '15'; Guid_{11997190-23841} '15'; ScreenModuleType ""
      on Guid_{11997190-21491}: SetTag("SelectedRack", 1); SetTag("SelectedSlot", 15); function_efd93a16("RackSlotData", 220, 150, -1, -1, 1)
      Guid_{11997190-21133} <- "WarehouseData_Rack1{15}"
   ScreenModuleView "RackSlot_18" at 262,315 size 44x36; Guid_{11997190-21654} '16'; Guid_{11997190-23841} '16'; ScreenModuleType ""
      on Guid_{11997190-21491}: SetTag("SelectedRack", 1); SetTag("SelectedSlot", 16); function_efd93a16("RackSlotData", 220, 150, -1, -1, 1)
      Guid_{11997190-21133} <- "WarehouseData_Rack1{16}"
   ScreenModuleView "RackSlot_19" at 212,315 size 44x36; Guid_{11997190-21654} '17'; Guid_{11997190-23841} '17'; ScreenModuleType ""
      on Guid_{11997190-21491}: SetTag("SelectedRack", 1); SetTag("SelectedSlot", 17); function_efd93a16("RackSlotData", 220, 150, -1, -1, 1)
      Guid_{11997190-21133} <- "WarehouseData_Rack1{17}"
   ScreenModuleView "RackSlot_20" at 162,315 size 44x36; Guid_{11997190-21654} '18'; Guid_{11997190-23841} '18'; ScreenModuleType ""
      on Guid_{11997190-21491}: SetTag("SelectedRack", 1); SetTag("SelectedSlot", 18); function_efd93a16("RackSlotData", 220, 150, -1, -1, 1)
      Guid_{11997190-21133} <- "WarehouseData_Rack1{18}"
   ScreenModuleView "RackSlot_21" at 562,270 size 44x36; Guid_{11997190-21654} '19'; Guid_{11997190-23841} '19'; ScreenModuleType ""
      on Guid_{11997190-21491}: SetTag("SelectedRack", 1); SetTag("SelectedSlot", 19); function_efd93a16("RackSlotData", 220, 150, -1, -1, 1)
      Guid_{11997190-21133} <- "WarehouseData_Rack1{19}"
   ScreenModuleView "RackSlot_22" at 512,270 size 44x36; Guid_{11997190-21654} '20'; Guid_{11997190-23841} '20'; ScreenModuleType ""
      on Guid_{11997190-21491}: SetTag("SelectedRack", 1); SetTag("SelectedSlot", 20); function_efd93a16("RackSlotData", 220, 150, -1, -1, 1)
      Guid_{11997190-21133} <- "WarehouseData_Rack1{20}"
   ScreenModuleView "RackSlot_23" at 462,270 size 44x36; Guid_{11997190-21654} '21'; Guid_{11997190-23841} '21'; ScreenModuleType ""
      on Guid_{11997190-21491}: SetTag("SelectedRack", 1); SetTag("SelectedSlot", 21); function_efd93a16("RackSlotData", 220, 150, -1, -1, 1)
      Guid_{11997190-21133} <- "WarehouseData_Rack1{21}"
   ScreenModuleView "RackSlot_24" at 412,270 size 44x36; Guid_{11997190-21654} '22'; Guid_{11997190-23841} '22'; ScreenModuleType ""
      on Guid_{11997190-21491}: SetTag("SelectedRack", 1); SetTag("SelectedSlot", 22); function_efd93a16("RackSlotData", 220, 150, -1, -1, 1)
      Guid_{11997190-21133} <- "WarehouseData_Rack1{22}"
   ScreenModuleView "RackSlot_25" at 362,270 size 44x36; Guid_{11997190-21654} '23'; Guid_{11997190-23841} '23'; ScreenModuleType ""
      on Guid_{11997190-21491}: SetTag("SelectedRack", 1); SetTag("SelectedSlot", 23); function_efd93a16("RackSlotData", 220, 150, -1, -1, 1)
      Guid_{11997190-21133} <- "WarehouseData_Rack1{23}"
   ScreenModuleView "RackSlot_26" at 312,270 size 44x36; Guid_{11997190-21654} '24'; Guid_{11997190-23841} '24'; ScreenModuleType ""
      on Guid_{11997190-21491}: SetTag("SelectedRack", 1); SetTag("SelectedSlot", 24); function_efd93a16("RackSlotData", 220, 150, -1, -1, 1)
      Guid_{11997190-21133} <- "WarehouseData_Rack1{24}"
   ScreenModuleView "RackSlot_27" at 262,270 size 44x36; Guid_{11997190-21654} '25'; Guid_{11997190-23841} '25'; ScreenModuleType ""
      on Guid_{11997190-21491}: SetTag("SelectedRack", 1); SetTag("SelectedSlot", 25); function_efd93a16("RackSlotData", 220, 150, -1, -1, 1)
      Guid_{11997190-21133} <- "WarehouseData_Rack1{25}"
   ScreenModuleView "RackSlot_28" at 212,270 size 44x36; Guid_{11997190-21654} '26'; Guid_{11997190-23841} '26'; ScreenModuleType ""
      on Guid_{11997190-21491}: SetTag("SelectedRack", 1); SetTag("SelectedSlot", 26); function_efd93a16("RackSlotData", 220, 150, -1, -1, 1)
      Guid_{11997190-21133} <- "WarehouseData_Rack1{26}"
   ScreenModuleView "RackSlot_29" at 162,270 size 44x36; Guid_{11997190-21654} '27'; Guid_{11997190-23841} '27'; ScreenModuleType ""
      on Guid_{11997190-21491}: SetTag("SelectedRack", 1); SetTag("SelectedSlot", 27); function_efd93a16("RackSlotData", 220, 150, -1, -1, 1)
      Guid_{11997190-21133} <- "WarehouseData_Rack1{27}"
   ScreenModuleView "RackSlot_30" at 562,225 size 44x36; Guid_{11997190-21654} '28'; Guid_{11997190-23841} '28'; ScreenModuleType ""
      on Guid_{11997190-21491}: SetTag("SelectedRack", 1); SetTag("SelectedSlot", 28); function_efd93a16("RackSlotData", 220, 150, -1, -1, 1)
      Guid_{11997190-21133} <- "WarehouseData_Rack1{28}"
   ScreenModuleView "RackSlot_31" at 512,225 size 44x36; Guid_{11997190-21654} '29'; Guid_{11997190-23841} '29'; ScreenModuleType ""
      on Guid_{11997190-21491}: SetTag("SelectedRack", 1); SetTag("SelectedSlot", 29); function_efd93a16("RackSlotData", 220, 150, -1, -1, 1)
      Guid_{11997190-21133} <- "WarehouseData_Rack1{29}"
   ScreenModuleView "RackSlot_32" at 462,225 size 44x36; Guid_{11997190-21654} '30'; Guid_{11997190-23841} '30'; ScreenModuleType ""
      on Guid_{11997190-21491}: SetTag("SelectedRack", 1); SetTag("SelectedSlot", 30); function_efd93a16("RackSlotData", 220, 150, -1, -1, 1)
      Guid_{11997190-21133} <- "WarehouseData_Rack1{30}"
   ScreenModuleView "RackSlot_33" at 412,225 size 44x36; Guid_{11997190-21654} '31'; Guid_{11997190-23841} '31'; ScreenModuleType ""
      on Guid_{11997190-21491}: SetTag("SelectedRack", 1); SetTag("SelectedSlot", 31); function_efd93a16("RackSlotData", 220, 150, -1, -1, 1)
      Guid_{11997190-21133} <- "WarehouseData_Rack1{31}"
   ScreenModuleView "RackSlot_34" at 362,225 size 44x36; Guid_{11997190-21654} '32'; Guid_{11997190-23841} '32'; ScreenModuleType ""
      on Guid_{11997190-21491}: SetTag("SelectedRack", 1); SetTag("SelectedSlot", 32); function_efd93a16("RackSlotData", 220, 150, -1, -1, 1)
      Guid_{11997190-21133} <- "WarehouseData_Rack1{32}"
   ScreenModuleView "RackSlot_35" at 312,225 size 44x36; Guid_{11997190-21654} '33'; Guid_{11997190-23841} '33'; ScreenModuleType ""
      on Guid_{11997190-21491}: SetTag("SelectedRack", 1); SetTag("SelectedSlot", 33); function_efd93a16("RackSlotData", 220, 150, -1, -1, 1)
      Guid_{11997190-21133} <- "WarehouseData_Rack1{33}"
   ScreenModuleView "RackSlot_36" at 262,225 size 44x36; Guid_{11997190-21654} '34'; Guid_{11997190-23841} '34'; ScreenModuleType ""
      on Guid_{11997190-21491}: SetTag("SelectedRack", 1); SetTag("SelectedSlot", 34); function_efd93a16("RackSlotData", 220, 150, -1, -1, 1)
      Guid_{11997190-21133} <- "WarehouseData_Rack1{34}"
   ScreenModuleView "RackSlot_37" at 212,225 size 44x36; Guid_{11997190-21654} '35'; Guid_{11997190-23841} '35'; ScreenModuleType ""
      on Guid_{11997190-21491}: SetTag("SelectedRack", 1); SetTag("SelectedSlot", 36); function_efd93a16("RackSlotData", 220, 150, -1, -1, 1)
      Guid_{11997190-21133} <- "WarehouseData_Rack1{35}"
   ScreenModuleView "RackSlot_38" at 162,225 size 44x36; Guid_{11997190-21654} '36'; Guid_{11997190-23841} '36'; ScreenModuleType ""
      on Guid_{11997190-21491}: SetTag("SelectedRack", 1); SetTag("SelectedSlot", 36); function_efd93a16("RackSlotData", 220, 150, -1, -1, 1)
      Guid_{11997190-21133} <- "WarehouseData_Rack1{36}"
   ScreenModuleView "RackSlot_39" at 562,180 size 44x36; Guid_{11997190-21654} '37'; Guid_{11997190-23841} '37'; ScreenModuleType ""
      on Guid_{11997190-21491}: SetTag("SelectedRack", 1); SetTag("SelectedSlot", 37); function_efd93a16("RackSlotData", 220, 150, -1, -1, 1)
      Guid_{11997190-21133} <- "WarehouseData_Rack1{37}"
   ScreenModuleView "RackSlot_40" at 512,180 size 44x36; Guid_{11997190-21654} '38'; Guid_{11997190-23841} '38'; ScreenModuleType ""
      on Guid_{11997190-21491}: SetTag("SelectedRack", 1); SetTag("SelectedSlot", 38); function_efd93a16("RackSlotData", 220, 150, -1, -1, 1)
      Guid_{11997190-21133} <- "WarehouseData_Rack1{38}"
   ScreenModuleView "RackSlot_41" at 462,180 size 44x36; Guid_{11997190-21654} '39'; Guid_{11997190-23841} '39'; ScreenModuleType ""
      on Guid_{11997190-21491}: SetTag("SelectedRack", 1); SetTag("SelectedSlot", 39); function_efd93a16("RackSlotData", 220, 150, -1, -1, 1)
      Guid_{11997190-21133} <- "WarehouseData_Rack1{39}"
   ScreenModuleView "RackSlot_42" at 412,180 size 44x36; Guid_{11997190-21654} '40'; Guid_{11997190-23841} '40'; ScreenModuleType ""
      on Guid_{11997190-21491}: SetTag("SelectedRack", 1); SetTag("SelectedSlot", 40); function_efd93a16("RackSlotData", 220, 150, -1, -1, 1)
      Guid_{11997190-21133} <- "WarehouseData_Rack1{40}"
   ScreenModuleView "RackSlot_43" at 362,180 size 44x36; Guid_{11997190-21654} '41'; Guid_{11997190-23841} '41'; ScreenModuleType ""
      on Guid_{11997190-21491}: SetTag("SelectedRack", 1); SetTag("SelectedSlot", 41); function_efd93a16("RackSlotData", 220, 150, -1, -1, 1)
      Guid_{11997190-21133} <- "WarehouseData_Rack1{41}"
   ScreenModuleView "RackSlot_44" at 312,180 size 44x36; Guid_{11997190-21654} '42'; Guid_{11997190-23841} '42'; ScreenModuleType ""
      on Guid_{11997190-21491}: SetTag("SelectedRack", 1); SetTag("SelectedSlot", 42); function_efd93a16("RackSlotData", 220, 150, -1, -1, 1)
      Guid_{11997190-21133} <- "WarehouseData_Rack1{42}"
   ScreenModuleView "RackSlot_45" at 262,180 size 44x36; Guid_{11997190-21654} '43'; Guid_{11997190-23841} '43'; ScreenModuleType ""
      on Guid_{11997190-21491}: SetTag("SelectedRack", 1); SetTag("SelectedSlot", 43); function_efd93a16("RackSlotData", 220, 150, -1, -1, 1)
      Guid_{11997190-21133} <- "WarehouseData_Rack1{43}"
   ScreenModuleView "RackSlot_46" at 212,180 size 44x36; Guid_{11997190-21654} '44'; Guid_{11997190-23841} '44'; ScreenModuleType ""
      on Guid_{11997190-21491}: SetTag("SelectedRack", 1); SetTag("SelectedSlot", 44); function_efd93a16("RackSlotData", 220, 150, -1, -1, 1)
      Guid_{11997190-21133} <- "WarehouseData_Rack1{44}"
   ScreenModuleView "RackSlot_47" at 162,180 size 44x36; Guid_{11997190-21654} '45'; Guid_{11997190-23841} '45'; ScreenModuleType ""
      on Guid_{11997190-21491}: SetTag("SelectedRack", 1); SetTag("SelectedSlot", 45); function_efd93a16("RackSlotData", 220, 150, -1, -1, 1)
      Guid_{11997190-21133} <- "WarehouseData_Rack1{45}"
   ScreenModuleView "RackSlot_48" at 562,135 size 44x36; Guid_{11997190-21654} '46'; Guid_{11997190-23841} '46'; ScreenModuleType ""
      on Guid_{11997190-21491}: SetTag("SelectedRack", 1); SetTag("SelectedSlot", 46); function_efd93a16("RackSlotData", 220, 150, -1, -1, 1)
      Guid_{11997190-21133} <- "WarehouseData_Rack1{46}"
   ScreenModuleView "RackSlot_49" at 512,135 size 44x36; Guid_{11997190-21654} '47'; Guid_{11997190-23841} '47'; ScreenModuleType ""
      on Guid_{11997190-21491}: SetTag("SelectedRack", 1); SetTag("SelectedSlot", 47); function_efd93a16("RackSlotData", 220, 150, -1, -1, 1)
      Guid_{11997190-21133} <- "WarehouseData_Rack1{47}"
   ScreenModuleView "RackSlot_50" at 462,135 size 44x36; Guid_{11997190-21654} '48'; Guid_{11997190-23841} '48'; ScreenModuleType ""
      on Guid_{11997190-21491}: SetTag("SelectedRack", 1); SetTag("SelectedSlot", 48); function_efd93a16("RackSlotData", 220, 150, -1, -1, 1)
      Guid_{11997190-21133} <- "WarehouseData_Rack1{48}"
   ScreenModuleView "RackSlot_51" at 412,135 size 44x36; Guid_{11997190-21654} '49'; Guid_{11997190-23841} '49'; ScreenModuleType ""
      on Guid_{11997190-21491}: SetTag("SelectedRack", 1); SetTag("SelectedSlot", 49); function_efd93a16("RackSlotData", 220, 150, -1, -1, 1)
      Guid_{11997190-21133} <- "WarehouseData_Rack1{49}"
   ScreenModuleView "RackSlot_52" at 362,135 size 44x36; Guid_{11997190-21654} '50'; Guid_{11997190-23841} '50'; ScreenModuleType ""
      on Guid_{11997190-21491}: SetTag("SelectedRack", 1); SetTag("SelectedSlot", 50); function_efd93a16("RackSlotData", 220, 150, -1, -1, 1)
      Guid_{11997190-21133} <- "WarehouseData_Rack1{50}"
   ScreenModuleView "RackSlot_53" at 312,135 size 44x36; Guid_{11997190-21654} '51'; Guid_{11997190-23841} '51'; ScreenModuleType ""
      on Guid_{11997190-21491}: SetTag("SelectedRack", 1); SetTag("SelectedSlot", 51); function_efd93a16("RackSlotData", 220, 150, -1, -1, 1)
      Guid_{11997190-21133} <- "WarehouseData_Rack1{51}"
   ScreenModuleView "RackSlot_54" at 262,135 size 44x36; Guid_{11997190-21654} '52'; Guid_{11997190-23841} '52'; ScreenModuleType ""
      on Guid_{11997190-21491}: SetTag("SelectedRack", 1); SetTag("SelectedSlot", 52); function_efd93a16("RackSlotData", 220, 150, -1, -1, 1)
      Guid_{11997190-21133} <- "WarehouseData_Rack1{52}"
   ScreenModuleView "RackSlot_55" at 212,135 size 44x36; Guid_{11997190-21654} '53'; Guid_{11997190-23841} '53'; ScreenModuleType ""
      on Guid_{11997190-21491}: SetTag("SelectedRack", 1); SetTag("SelectedSlot", 53); function_efd93a16("RackSlotData", 220, 150, -1, -1, 1)
      Guid_{11997190-21133} <- "WarehouseData_Rack1{53}"
   ScreenModuleView "RackSlot_56" at 162,135 size 44x36; Guid_{11997190-21654} '54'; Guid_{11997190-23841} '54'; ScreenModuleType ""
      on Guid_{11997190-21491}: SetTag("SelectedRack", 1); SetTag("SelectedSlot", 54); function_efd93a16("RackSlotData", 220, 150, -1, -1, 1)
      Guid_{11997190-21133} <- "WarehouseData_Rack1{54}"
   TextField "Text field_1" at 17,171 size 106x22; Text 'Crane Status:'
   TextField "Text field_2" at 17,360 size 113x22; Text 'Both racks full'
      Visibility <- "RacksFull"
   TextField "Text field_4" at 15,121 size 15x22; Text 'Text'
   TextField "Text field_3" at 17,193 size 70x18; Text 'Text'
   TextField "Text field_5" at 17,261 size 119x22; Text 'Occupied slots:'
   TextField "Text field_6" at 36,283 size 28x18; Text '/ 54'
   TextField "Text field_7" at 17,283 size 29x18; Text 'Text'
   Button "Button_3" at 17,104 size 54x39; TextOff 'START'
      on Press: SetBit("StartCmd")
      on Release: ResetBit("StartCmd")
   Button "Button_4" at 80,104 size 54x39; TextOff 'STOP'
      on Press: SetBit("StopCmd")
      on Release: ResetBit("StopCmd")

PopupScreen "RackSlotData" 240x200
   TextField "Text field_1" at 18,26 size 74x22; Text 'Pallet Id:'
   TextField "Text field_2" at 64,87 size 108x22; Text 'Storage Date:'
   TextField "Text field_3" at 18,48 size 58x22; Text 'Status:'
   Button "Button_1" at 15,153 size 96x32; TextOff 'Retrieve'
      on Click: function_efd93a16("ConfirmRequest", 220, 150, 1, -1, 1)
      ObjectEnable <- "Status"
      Appearance <- "Status"
   TextField "Text field_4" at 156,26 size 50x22; Text 'Text'
   TextField "Text field_5" at 15,109 size 213x22; Text 'Text'
   TextField "Text field_6" at 156,48 size 76x22; Text 'Text'
   Button "Button_2" at 132,153 size 96x32; TextOff 'Close'
      on Click: function_efd93a16("RackSlotData", 0, 0, 0, -1, 1)

PopupScreen "ConfirmRequest" 240x100
   Button "Button_2" at 134,64 size 87x24; TextOff 'No'
      on Click: function_efd93a16("ConfirmRequest", 0, 0, 0, -1, 1)
   Button "Button_1" at 20,64 size 87x24; TextOff 'Yes'
      on Press: SetBit("RetrievePallet")
      on Release: ResetBit("RetrievePallet"); function_efd93a16("ConfirmRequest", 0, 0, 0, -1, 1)
   TextField "Text field_1" at 20,7 size 201x40; Text 'Do you want to send a pallet retrieval request?'

